(* IEC 61131-3 sources: daoli-st-library/DL_Device (part 16) *)

(* ---- FB_DL_CleanRoomRhTrim.st ---- *)
(*
  FB_DL_CleanRoomRhTrim  —  洁净室加湿阀脉冲微调（RH 偏差 + 最小开度保护） / Clean-room humidifier pulse trim with RH deviation and minimum-opening protection
  分类 Category : DL_Device
  版本 Version  : 1.0.0
  来源 Source   : t1-2-oscat-building — 楼宇洁净室湿度控制族深化
  溯源 Origin   : 道莅 clean-room 实现；脉宽调制加湿（PWM 占空比 + 最小开度 + 高限停加湿）为公开洁净室湿度算法，未复制任何源码行
  功能 Function : 1) 每个脉冲周期起始重算占空比：duty = fKpPctPerPct × (fRhSpPct - fRhPct)，
                  钳制到 [0.0, 100.0]；
                  2) 最小开度保护：fRhPct 低于 fRhLoPct 时 duty 取 max(duty, fMinOpenPct)；
                  3) 高限停加湿：fRhPct 高于 fRhHiPct 时 duty 强制 0（防过湿）；
                  4) 脉宽：开阀时长 = duty × tPeriod / 100.0（除数常量 100.0），关阀时长 = 周期余量；
                  5) 故障级单码 052B / 信息级 0431 = 脉冲周期完成沿（每周期单拍）。
  接口 Interface: 输入 RH 设定/实测/上下限/增益/最小开度/周期；输出阀指令与占空比镜像
  边界 Boundary : ① 组态闸：tPeriod <= T#0S、fMinOpenPct 不在 [0,100]、fKpPctPerPct <= 0.0、
                  fRhHiPct <= fRhLoPct、fRhSpPct 不在 [0,100] → 052B 锁存；
                  ② RH 非有限（NaN 自反 + Inf 差值自减）→ 052B 锁存，阀指令强制关断；
                  ③ 占空比开阀时长按实数乘除后转 TIME，转换前钳制到 [0, tPeriod] 防越界；
                  ④ 两个 TON 段 0 无条件周期调用，IN 由相位/占空比派生，相内自动复位 ET；
                  ⑤ 故障相迁出唯一路径 = bReset 上升沿；⑥ 零全局耦合（无 GVL / %I %Q %M）。
  依赖 Depends  : Standard.library（TON / R_TRIG）
  码表 Error codes（Device 分段见下，故障窗口 052B / 信息窗口 0431）:
    16#0003_052B 故障级：加湿脉冲故障总码（组态非法 / RH 非有限），锁存至 bReset 上升沿；
                 归因见 eCause，不新增码位（派单硬约束单码）
    16#0003_0431 信息级：脉冲周期完成沿（占空比重算单拍）
    分段理由：段 0003 故障带 03A0~03FF 于 R42 用尽，启用 05xx 副带续编，避开 0590~0599 判错位段。
  修订历史 Revision :
    2026-11-19  v1.0.0  R43 首版（批次 3 · 序号 15）
*)

TYPE E_DL_CrhState :
(
    eIdle  := 0,      // 未使能：阀关 / Idle, valve closed
    ePulse := 10,     // 脉冲调制中（开/关按时长切换） / Pulse modulation
    eFault := 90      // 故障锁存相（阀强制关） / Fault latched, valve forced closed
);
END_TYPE

TYPE E_DL_CrhCause :
(
    eNone       := 0, // 无故障成因 / No cause
    eCfgIllegal := 1, // 组态非法 / Illegal configuration
    eNonFinite  := 2  // RH 非有限 / Non-finite RH
);
END_TYPE

FUNCTION_BLOCK FB_DL_CleanRoomRhTrim
VAR_INPUT
    fRhSpPct      : REAL := 45.0;      // RH 设定 [%]，域 [0,100] / RH setpoint
    fRhPct        : REAL := 0.0;       // RH 实测 [%] / Measured RH
    fRhLoPct      : REAL := 40.0;      // 低限（触发最小开度） [%] / Low limit for minimum opening
    fRhHiPct      : REAL := 55.0;      // 高限（停加湿） [%] / High limit stopping humidification
    fKpPctPerPct  : REAL := 8.0;       // 比例增益 [%/ %]，域 > 0 / Proportional gain
    fMinOpenPct   : REAL := 10.0;      // 最小开度 [%]，域 [0,100] / Minimum opening
    tPeriod       : TIME := T#10S;     // 脉冲周期 [ms]，域 > 0 / Pulse period
    bEnable       : BOOL := FALSE;     // 加湿使能（电平）[-] / Humidification enable
    bReset        : BOOL := FALSE;     // 复位命令，上升沿清故障 [-] / Reset edge
END_VAR
VAR_OUTPUT
    eState        : E_DL_CrhState;     // 状态出口，段 6 单点映射 / State outlet
    eCause        : E_DL_CrhCause;     // 故障成因出口（R190） / Fault cause outlet
    bHumValve     : BOOL;              // 加湿阀指令 [-] / Humidifier valve command
    fDutyPct      : REAL;              // 占空比镜像 [%] / Duty mirror
    bMinOpen      : BOOL;              // 最小开度生效镜像 [-] / Minimum opening active
    bCycleDone    : BOOL;              // 脉冲周期完成标志 [-] / Pulse period done flag
    bError        : BOOL;              // 故障锁存标志 [-] / Fault latch flag
    nErrId        : UDINT;             // 事件码，0 = 无事件 / Event code
END_VAR
VAR
    _eState       : E_DL_CrhState := E_DL_CrhState.eIdle;   // 内部相位（CASE 唯一写入目标） / Internal phase
    _eCause       : E_DL_CrhCause := E_DL_CrhCause.eNone;   // 故障成因锁存（锁存量） / Latched cause
    tonOn         : TON;               // 开阀时长计时，每周期无条件调用 / Valve-on timer
    tonOff        : TON;               // 关阀时长计时，每周期无条件调用 / Valve-off timer
    rtReset       : R_TRIG;            // 复位沿实例，每周期无条件调用 / Reset edge
    _fDutyPct     : REAL;              // 占空比保持量（本周期内恒定） / Duty held for the period
    _fOnMs        : REAL;              // 本周期开阀时长 [ms]（钳制后） / On-time in ms
    _fOffMs       : REAL;              // 本周期关阀时长 [ms] / Off-time in ms
    _bOnPhase     : BOOL;              // 当前处于开阀段（内部相位标志） / In on-segment flag
    _bMinOpenOn   : BOOL;              // 最小开度生效当拍量 [-] / Minimum opening flag
    _bNonFin      : BOOL;              // RH 非有限当拍量 [-] / Non-finite RH
    _bCfgBad      : BOOL;              // 组态非法当拍量 [-] / Config illegal
    _bFault       : BOOL;              // 故障锁存位（锁存量） / Latched fault bit
    _uFault       : UDINT;             // 故障码锁存（锁存量） / Latched fault code
    _uInfo        : UDINT;             // 信息码，每拍重算 / Transient info code
END_VAR

(* —— 段 0：沿实例与定时器无条件周期刷新 + 当拍量判据 —— *)
_bNonFin := (fRhPct <> fRhPct) OR (fRhSpPct <> fRhSpPct)
         OR ((fRhPct - fRhPct) <> (fRhPct - fRhPct))
         OR ((fRhSpPct - fRhSpPct) <> (fRhSpPct - fRhSpPct));                 // NaN 自反 + Inf 差值自减 / NaN and Inf
_bCfgBad := (tPeriod <= T#0S) OR (fKpPctPerPct <= 0.0) OR (fRhHiPct <= fRhLoPct)
            OR (fMinOpenPct < 0.0) OR (fMinOpenPct > 100.0)
            OR (fRhSpPct < 0.0) OR (fRhSpPct > 100.0);                        // 组态非法当拍量 / Config illegal
rtReset(CLK := bReset);                                                       // 复位沿，每拍必调 / Reset edge
tonOn(IN := (_bOnPhase AND (_eState = E_DL_CrhState.ePulse)), PT := REAL_TO_TIME(_fOnMs));    // 开阀计时（实数时长转 TIME） / On timer
tonOff(IN := (NOT _bOnPhase) AND (_eState = E_DL_CrhState.ePulse), PT := REAL_TO_TIME(_fOffMs));  // 关阀计时 / Off timer

(* —— 段 1：单拍量预清零（锁存量与占空比保持量不入清单） —— *)
_uInfo := 16#0000_0000;            // 信息码每拍重算 / Info recomputed
bHumValve := FALSE;                // 阀指令缺省关 / Valve command default closed
fDutyPct := 0.0;                   // 占空比出口缺省 0 / Duty default
bMinOpen := FALSE;                 // 最小开度镜像缺省 FALSE / Minimum opening default
bCycleDone := FALSE;               // 周期完成标志缺省 FALSE / Period done default
nErrId := 16#0000_0000;            // 事件码缺省无事件 / Event code default

(* —— 段 2：复位沿 + 组态域闸 —— *)
IF rtReset.Q THEN                              // rtReset.Q = 当拍量 / current scan
    _bFault := FALSE;                          // 清故障锁存位（锁存量） / Clear fault latch
    _uFault := 16#0000_0000;                   // 清故障锁存码（锁存量） / Clear fault code
    _eCause := E_DL_CrhCause.eNone;            // 清成因（锁存量） / Clear cause
    _fDutyPct := 0.0;                          // 清占空比保持量 / Clear duty
    _bOnPhase := FALSE;                        // 清开阀段标志 / Clear on-segment
    IF _eState = E_DL_CrhState.eFault THEN
        _eState := E_DL_CrhState.eIdle;        // 故障相迁出：回未使能 / Fault exit to idle
    END_IF
END_IF
IF _bCfgBad THEN                               // 组态域闸 / Config gate
    _uFault := 16#0003_052B;                   // 故障级：加湿脉冲故障总码（05xx 副带） / Device fault code
    _eCause := E_DL_CrhCause.eCfgIllegal;      // 归因：组态非法 / Cause: illegal config
    _bFault := TRUE;                           // 标志与码位配对（R45） / Flag paired with code
END_IF
IF (NOT _bFault) AND _bNonFin THEN             // 非有限锁存 / Non-finite latch
    _uFault := 16#0003_052B;
    _eCause := E_DL_CrhCause.eNonFinite;       // 归因：非有限 / Cause: non-finite
    _bFault := TRUE;
END_IF

(* —— 段 3：占空比重算（周期边界 = 关阀段结束或首次进入） —— *)
IF (NOT _bFault) AND (_eState = E_DL_CrhState.ePulse) AND tonOff.Q THEN
    _fDutyPct := fKpPctPerPct * (fRhSpPct - fRhPct);                  // 比例占空比 [%] / Proportional duty
    IF fRhPct < fRhLoPct THEN                                        // 低限：最小开度保护 / Low limit protection
        IF _fDutyPct < fMinOpenPct THEN
            _fDutyPct := fMinOpenPct;                                // 抬到最小开度 / Raise to minimum
            _bMinOpenOn := TRUE;
        END_IF
    END_IF
    IF fRhPct > fRhHiPct THEN                                        // 高限：停加湿 / High limit stops humidification
        _fDutyPct := 0.0;
        _bMinOpenOn := FALSE;
    END_IF
    IF _fDutyPct < 0.0 THEN                                          // 占空比下限钳制 / Duty low clamp
        _fDutyPct := 0.0;
    ELSIF _fDutyPct > 100.0 THEN                                     // 占空比上限钳制 / Duty high clamp
        _fDutyPct := 100.0;
    END_IF
    _fOnMs := _fDutyPct / 100.0 * TIME_TO_REAL(tPeriod);             // 开阀时长 [ms]（除常量 100.0） / On-time
    IF _fOnMs < 0.0 THEN                                             // 时长下限钳制（防负数） / On-time low clamp
        _fOnMs := 0.0;
    ELSIF _fOnMs > TIME_TO_REAL(tPeriod) THEN                        // 时长上限钳制（不越周期） / On-time high clamp
        _fOnMs := TIME_TO_REAL(tPeriod);
    END_IF
    _fOffMs := TIME_TO_REAL(tPeriod) - _fOnMs;                       // 关阀时长 = 周期余量 / Off-time remainder
    _uInfo := 16#0003_0431;                                          // 信息级：脉冲周期完成沿 / Info: period done edge
END_IF

(* —— 段 4：故障解除式（R240；全当拍量）：rtReset.Q / NOT _bCfgBad / NOT _bNonFin —— *)
IF rtReset.Q AND (NOT _bCfgBad) AND (NOT _bNonFin) THEN
    _bFault := FALSE;                          // 清故障锁存位（锁存量） / Clear fault latch
    _uFault := 16#0000_0000;                   // 清故障锁存码（锁存量） / Clear fault code
    _eCause := E_DL_CrhCause.eNone;            // 清成因（锁存量） / Clear cause
END_IF

(* —— 段 4A：故障锁存相位迁移闸（阀强制关） —— *)
IF _bFault AND (_eState <> E_DL_CrhState.eFault) THEN
    _eState := E_DL_CrhState.eFault;           // 锁存即入故障相 / Latch enters fault phase
END_IF

(* —— 段 5：相位机（CASE 全覆盖 + ELSE 兜底） —— *)
CASE _eState OF

E_DL_CrhState.eIdle:
    IF bEnable AND (NOT _bFault) THEN          // 使能条件 / Enable gate
        _fDutyPct := 0.0;                      // 起始占空比 0 / Start duty zero
        _fOnMs := 0.0;                         // 起始开阀时长 0 / Start on-time zero
        _fOffMs := TIME_TO_REAL(tPeriod);      // 起始关阀时长 = 整周期 / Start off-time full period
        _bOnPhase := FALSE;                    // 从关阀段起步 / Start in off-segment
        _eState := E_DL_CrhState.ePulse;       // 进脉冲相 / Enter pulse
    END_IF

E_DL_CrhState.ePulse:
    IF _bOnPhase THEN                          // 开阀段 / On-segment
        bHumValve := TRUE;                     // 阀开 / Valve open
        IF tonOn.Q THEN                        // 开阀到时 / On-time elapsed
            _bOnPhase := FALSE;                // 转关阀段 / Switch to off-segment
        END_IF
    ELSE
        bHumValve := FALSE;                    // 阀关 / Valve closed
        IF (_fOnMs > 0.0) AND tonOff.Q THEN    // 关阀到时且有开阀时长 / Off-time elapsed with on-time
            _bOnPhase := TRUE;                 // 转开阀段 / Switch to on-segment
        ELSIF (_fOnMs <= 0.0) AND tonOff.Q THEN
            ;                                  // 零占空比：保持关阀（周期照常走完） / Zero duty keeps valve closed
            _bOnPhase := FALSE;
        END_IF
    END_IF
    IF NOT bEnable THEN                        // 撤使能：阀关，回未使能 / Disable closes valve
        _bOnPhase := FALSE;
        _eState := E_DL_CrhState.eIdle;
    END_IF

E_DL_CrhState.eFault:
    ;                                          // 故障相：阀强制关，仅段 4 复位沿可迁出 / Valve closed, reset only

ELSE
    _uFault := 16#0003_052B;                   // 故障级：非法相位兜底（归并总码） / Illegal phase fallback
    _eCause := E_DL_CrhCause.eCfgIllegal;      // 归因：相位非法归并组态 / Cause: phase illegal
    _bFault := TRUE;
    _eState := E_DL_CrhState.eFault;           // 强制回故障相 / Force fault phase

END_CASE

(* —— 段 6：出口单点映射（名实同源；故障相阀强制关断） —— *)
IF _bFault THEN
    bHumValve := FALSE;                        // 故障相阀强制关（安全侧） / Valve forced closed
    nErrId := _uFault;                         // 故障锁存码回放 / Replay latched code
    fDutyPct := 0.0;                           // 故障相占空比强制 0 / Duty forced zero
    bMinOpen := FALSE;                         // 故障相最小开度镜像强制 FALSE / Minimum opening forced false
ELSE
    nErrId := _uInfo;                          // 信息码 / Transient info
    fDutyPct := _fDutyPct;                     // 占空比镜像 / Duty mirror
    bMinOpen := _bMinOpenOn;                   // 最小开度镜像 / Minimum opening mirror
END_IF
bCycleDone := (_eState = E_DL_CrhState.ePulse) AND tonOff.Q;   // 周期完成标志（当拍量） / Period done flag
bError := _bFault;                             // 故障标志同源 / Flag from latch
eState := _eState;                             // 状态出口 / State outlet
eCause := _eCause;                             // 成因出口 / Cause outlet

END_FUNCTION_BLOCK

(* ---- FB_DL_CncLoadUnloadSeq.st ---- *)
(*
  DL Factory R84 | FB_DL_CncLoadUnloadSeq
  功能：机床上下料八相时序状态机，逐相超时置故障码并锁存至复位沿
  开源溯源：无（clean-room 自研，依据公开工艺公式，来源=行业通用公式，许可证=MIT，借鉴点=公式结构）
  规则：R1-R16 全遵守
*)
TYPE E_DL_CncUsState :
(
    eIdle := 0, // 空闲待启动 [-] / idle, waiting for start [-]
    eDoorOpen := 1, // 开门相 [-] / door opening phase [-]
    eClampOpen := 2, // 夹具松开相 [-] / clamp opening phase [-]
    ePartLoad := 3, // 上料相 [-] / part loading phase [-]
    eClampClose := 4, // 夹具夹紧相 [-] / clamp closing phase [-]
    eDoorClose := 5, // 关门相 [-] / door closing phase [-]
    eCycleStart := 6, // 加工启动相 [-] / cycle start phase [-]
    eDone := 7, // 完成相 [-] / done phase [-]
    eFault := 8 // 故障锁存相 [-] / fault latched phase [-]
) := eIdle;
END_TYPE

FUNCTION_BLOCK FB_DL_CncLoadUnloadSeq
VAR_INPUT
    xStart : BOOL; // 启动按钮 [-] / start pushbutton [-]
    xReset : BOOL; // 复位按钮（上升沿清故障码） [-] / reset pushbutton [-]
    xDoorOpened : BOOL; // 门开到位反馈 [-] / door open limit [-]
    xDoorClosed : BOOL; // 门关到位反馈 [-] / door closed limit [-]
    xClampOpened : BOOL; // 夹具松开到位反馈 [-] / clamp open limit [-]
    xClampClosed : BOOL; // 夹具夹紧到位反馈 [-] / clamp closed limit [-]
    xPartPresent : BOOL; // 工件在位检测 [-] / part present sensor [-]
    xCycleAllowed : BOOL; // 加工许可互锁（外部给定） [-] / cycle permit interlock [-]
    xCycleDone : BOOL; // 加工完成反馈 [-] / cycle finished feedback [-]
    tPhaseLimit : TIME := T#10S; // 单相超时门限 [s] / per phase timeout limit [s]
END_VAR
VAR_OUTPUT
    eState : E_DL_CncUsState; // 当前时序状态 [-] / current sequence state [-]
    iErrCode : INT; // 故障码 0=正常，101~106=逐相超时，201=非法相位 [-] / error code [-]
    xBusy : BOOL; // 时序执行中 [-] / sequence busy [-]
    xDone : BOOL; // 完成单拍脉冲 [-] / done one-shot pulse [-]
END_VAR
VAR
    rtStart : R_TRIG; // 启动上升沿实例 [-] / start rising edge instance [-]
    rtReset : R_TRIG; // 复位上升沿实例 [-] / reset rising edge instance [-]
    tonPhase : TON; // 相超时定时器（全相共用） [-] / shared phase timeout timer [-]
    xTimerRun : BOOL; // 定时器运行使能 [-] / timer run enable [-]
    tLimit : TIME; // 当前相超时设定 [s] / current phase timeout preset [s]
    xTimeout : BOOL; // 本拍超时标志 [-] / timeout flag of this scan [-]
    xDoneInt : BOOL; // 完成内部锁存位 [-] / internal done latch [-]
    xDonePrev : BOOL; // 完成前拍快照 [-] / done previous scan snapshot [-]
    _eState : E_DL_CncUsState := E_DL_CncUsState.eIdle; // 内部相位（CASE 唯一写目标） [-] / internal phase [-]
    _ePrev : E_DL_CncUsState := E_DL_CncUsState.eIdle; // 相位前拍快照（供自复位判沿） [-] / previous phase snapshot [-]
    xPhaseChg : BOOL; // 相位切换当拍标志 [-] / phase change flag of this scan [-]
    _iErr : INT; // 故障码内部锁存 [-] / latched error code [-]
END_VAR

// 段 0｜边沿实例无条件周期刷新（R7）
rtStart(CLK := xStart); // 启动沿每拍必调 [-] / start edge called every scan [-]
rtReset(CLK := xReset); // 复位沿每拍必调 [-] / reset edge called every scan [-]

// 段 1｜按相位选超时预设（必须在定时器调用之前完成）
CASE _eState OF
    E_DL_CncUsState.eIdle: tLimit := T#0S; // 空闲不计时 [s] / no timing in idle [s]
    E_DL_CncUsState.eDone: tLimit := T#0S; // 完成不计时 [s] / no timing in done [s]
    E_DL_CncUsState.eFault: tLimit := T#0S; // 故障不计时 [s] / no timing in fault [s]
ELSE
    tLimit := tPhaseLimit; // 其余工作相按门限计时 [s] / working phases use the limit [s]
END_CASE

// 段 2｜定时器无条件周期刷新（CASE 之外，无 IF 包裹；换相即自复位，R7/R188）
xPhaseChg := _eState <> _ePrev; // 相位切换沿 [-] / phase change edge [-]
xTimerRun := (((_eState <> E_DL_CncUsState.eIdle) AND (_eState <> E_DL_CncUsState.eDone)) AND (_eState <> E_DL_CncUsState.eFault)) AND NOT xPhaseChg; // 工作相定时使能，换相当拍拉低以复位计时 [-] / timing enable, dropped on a phase change to restart [-]
tonPhase(IN := xTimerRun, PT := tLimit); // 无条件刷新 [-] / unconditional refresh [-]
xTimeout := tonPhase.Q; // 本拍超时判定 [-] / timeout verdict of this scan [-]
_ePrev := _eState; // 相位快照在定时器之后更新（本拍迁移下一拍生效） [-] / phase snapshot updated after the timer call [-]

// 段 3｜复位沿：清单为故障码 + 内部锁存 + 相位，不含 Prev/Acc 保持量（R189）
IF rtReset.Q THEN
    _iErr := 0; // 清故障码 [-] / clear error code [-]
    xDoneInt := FALSE; // 清完成锁存 [-] / clear done latch [-]
    _eState := E_DL_CncUsState.eIdle; // 回空闲相 [-] / back to idle [-]
END_IF

// 段 4｜主状态机（合法事件优先于超时迁移，R275）
CASE _eState OF
    E_DL_CncUsState.eIdle: // 空闲相 [-] / idle [-]
        xDoneInt := FALSE; // 空闲清完成锁存 [-] / clear done latch in idle [-]
        IF rtStart.Q THEN
            _eState := E_DL_CncUsState.eDoorOpen; // 启动沿开安全门 [-] / start edge opens the door [-]
        END_IF
    E_DL_CncUsState.eDoorOpen: // 开门相 [-] / door opening [-]
        IF xDoorOpened THEN
            _eState := E_DL_CncUsState.eClampOpen; // 门开到位转松夹 [-] / door open leads to clamp open [-]
        ELSIF xTimeout THEN
            _iErr := 101; _eState := E_DL_CncUsState.eFault; // 开门超时 [-] / door open timeout [-]
        END_IF
    E_DL_CncUsState.eClampOpen: // 松夹相 [-] / clamp opening [-]
        IF xClampOpened THEN
            _eState := E_DL_CncUsState.ePartLoad; // 松夹到位转上料 [-] / clamp open leads to loading [-]
        ELSIF xTimeout THEN
            _iErr := 102; _eState := E_DL_CncUsState.eFault; // 松夹超时 [-] / clamp open timeout [-]
        END_IF
    E_DL_CncUsState.ePartLoad: // 上料相 [-] / part loading [-]
        IF xPartPresent AND NOT xTimeout THEN
            _eState := E_DL_CncUsState.eClampClose; // 工件在位转夹紧（带超时复检） [-] / part present leads to clamp close [-]
        ELSIF xTimeout THEN
            _iErr := 103; _eState := E_DL_CncUsState.eFault; // 上料超时（工件未到位） [-] / loading timeout [-]
        END_IF
    E_DL_CncUsState.eClampClose: // 夹紧相 [-] / clamp closing [-]
        IF xClampClosed THEN
            _eState := E_DL_CncUsState.eDoorClose; // 夹紧到位转关门 [-] / clamp closed leads to door close [-]
        ELSIF xTimeout THEN
            _iErr := 104; _eState := E_DL_CncUsState.eFault; // 夹紧超时 [-] / clamp close timeout [-]
        END_IF
    E_DL_CncUsState.eDoorClose: // 关门相 [-] / door closing [-]
        IF xDoorClosed THEN
            _eState := E_DL_CncUsState.eCycleStart; // 关门到位转加工启动 [-] / door closed leads to cycle start [-]
        ELSIF xTimeout THEN
            _iErr := 105; _eState := E_DL_CncUsState.eFault; // 关门超时 [-] / door close timeout [-]
        END_IF
    E_DL_CncUsState.eCycleStart: // 加工启动相（执行类安全相，入相全量复检） [-] / cycle start [-]
        IF xCycleDone THEN
            _eState := E_DL_CncUsState.eDone; // 加工完成转完成相 [-] / cycle done leads to done [-]
        ELSIF NOT (xCycleAllowed AND xDoorClosed) THEN
            _iErr := 106; _eState := E_DL_CncUsState.eFault; // 许可消失即故障（不空等） [-] / permit lost becomes fault [-]
        ELSIF xTimeout THEN
            _iErr := 106; _eState := E_DL_CncUsState.eFault; // 加工未完成超时 [-] / cycle start timeout [-]
        END_IF
    E_DL_CncUsState.eDone: // 完成相 [-] / done [-]
        xDoneInt := TRUE; // 置完成锁存（出口统一映射单拍） [-] / raise done latch [-]
        IF NOT xStart THEN
            _eState := E_DL_CncUsState.eIdle; // 松开启动即回空闲 [-] / start released returns to idle [-]
        END_IF
    E_DL_CncUsState.eFault: // 故障相：码值锁存回放，仅复位沿出 [-] / fault, exit only on reset edge [-]
        ; // 锁存回放，不按当下输入重新推断（R28） [-] / replay the latch only [-]
ELSE
    _iErr := 201; _eState := E_DL_CncUsState.eFault; // 非法相位兜底 [-] / illegal phase fallback [-]
END_CASE

// 段 5｜出口映射（名实双出口，同源赋值）
eState := _eState; // 状态出口 [-] / state outlet [-]
iErrCode := _iErr; // 故障码出口（锁存值） [-] / error code outlet [-]
xBusy := ((_eState <> E_DL_CncUsState.eIdle) AND (_eState <> E_DL_CncUsState.eDone)) AND (_eState <> E_DL_CncUsState.eFault); // 忙 = 工作相镜像 [-] / busy mirrors a working phase [-]
xDone := xDoneInt AND NOT xDonePrev; // 完成单拍（内部锁存 → 出口映射） [-] / done one-shot [-]
xDonePrev := xDoneInt; // 本拍快照供下拍比较 [-] / snapshot for the next scan [-]
END_FUNCTION_BLOCK

(* ---- FB_DL_CncToolWearCompLoop.st ---- *)
(*
  DL Factory R84 | FB_DL_CncToolWearCompLoop
  功能：CNC 刀具后刀面磨损量 VB 在线估计与刀补闭环：按切削路程三段线性磨损曲线出 VB 原值，按切削比能调制滤波增益做一阶指数平滑得 VB 估计，超补偿门限按增量限幅出刀补，超寿命锁存换刀请求。
  开源溯源：无（clean-room 自研，依据公开工艺公式与安全设计惯例，来源=行业通用公式+工程实践，许可证=MIT，借鉴点=公式结构与联锁分层）
  规则：R1-R16 全遵守
  ------------------------------------------------------------------
  分类 DL_Device ｜ 复杂度 cx4 ｜ 版本 v1.0.0 ｜ 平台 纯 IEC 61131-3（LREAL、ENUM、CASE）
  边界一：只出刀补增量与换刀请求，不驱动伺服轴、不写 CNC 刀补表（落表由上层 PRG 执行，属主边界）。
  边界二：磨损曲线为三段线性——初期占额定寿命路程 0.15 段、占磨损余量 0.30 份；稳态占 0.70 段、占 0.55 份；
          急剧占余下 0.15 段、占余下 0.15 份；三段积分在路程等于额定寿命处恰等于 VB 限值（量纲自检见下）。
  边界三：切削路程按「进给率 × 切削时长增量」积分，时长增量取 fCutTimeS 的上拍快照差分（R45 ②）；
          负增量判零、超大跳变钳到 1 秒，防掉电恢复的时钟跳变伪造路程。
  边界四：工艺代理常量——DL_CNC_AP_MM 与 DL_CNC_AE_MM 为名义切深与切宽代理值（本件无切深切宽引脚）；
          代理值是名义切深切宽、覆盖常规铣削 0.2~3 mm 切深与 4~20 mm 切宽区间、区间外的重型切槽工况由上层
          按实际切深切宽折算 fKcNmm2 后下发（R95 三句齐备，代理假设挂编译验证债）。
  边界五：无效拍语义——功率或转速为零、或任一浮点入参非有限 → xValid 出假、相位保持、刀补增量出零；
          不推进滤波、不累加路程（不除零、不外推）。
  边界六：换刀请求 xChangeReq 为锁存式，唯一解除路径为 bReset 上升沿（R188）；xAlarm 为电平式跟随相位。
  量纲自检：VB [mm]＝斜率 [mm/m] × 路程 [m]；斜率一 ＝ VB限值 × 0.30 ÷（额定寿命 × 0.15）[mm/m]；
          路程增量 [m]＝进给 [mm/min] × 时长增量 [s] ÷ 60 [s/min] × 0.001 [m/mm]；
          切削功率 [kW]＝Kc [N/mm²] × 切除率 [mm³/s] ÷ 1000 [W/kW]；
          切除率 [mm³/s]＝进给 [mm/s] × 切深 [mm] × 切宽 [mm]；刀补 [µm]＝VB [mm] × 1000 [µm/mm]。
  码表：本件全部码位为信息级（2601 非法相位、2602 组态越域、2603 入参非有限、2604 转速或功率为零）；
        信息级码每拍重算且不置 bError；故障级语义由 xChangeReq 锁存位承担，故本件无 bError 出口（R187）。
  输出契约：fCompUm 为本次刀补增量 [µm]（限幅 ±50，非补偿相出 0 不保持）；fCompAccUm 为累计刀补 [µm]（0~200 单向）；
          fVbEst 为滤波后估计 [mm]；fVbRaw 为曲线原值 [mm]；iErrCode 信息级，非零时 xValid 恒假。
  修订记录：2026-11-24 v1.0.0 R84 首版（批 R84 · 序号 41）
*)

TYPE E_DL_CncWearState :
(
    eIdle       := 0,  // 空闲：等使能与切削条件 / idle, waiting for the enable and the cutting condition
    eLearn      := 10, // 学习：累加路程并收敛 VB 滤波 / learning, accumulate the path and settle the filter
    eCompensate := 20, // 补偿：VB 超补偿门限，按增量出刀补 / compensating, the wear passed the trigger threshold
    eAlarm      := 30, // 报警：VB 超报警门限，继续补偿并报警 / alarm, the wear passed the alarm threshold
    eChangeReq  := 40  // 换刀请求：VB 超寿命，锁存至复位沿 / change request, the wear passed the life limit and is latched
);
END_TYPE

TYPE E_DL_CncWearCause :
(
    eNone      := 0, // 无成因 / no cause
    ePhaseBad  := 1, // 非法相位（信息级 2601）/ illegal phase, info grade 2601
    eCfgBad    := 2, // 组态越域（信息级 2602）/ the configuration is out of its domain, info grade 2602
    eNotFinite := 3, // 入参非有限（信息级 2603）/ a non-finite input, info grade 2603
    eSpeedZero := 4  // 转速或功率为零（信息级 2604）/ the speed or the power is zero, info grade 2604
);
END_TYPE

FUNCTION_BLOCK FB_DL_CncToolWearCompLoop
VAR CONSTANT
    DL_CNC_PH1_FRAC   : LREAL := 0.15;    // 初期磨损段占额定寿命的路程分数 [-] / the initial wear path fraction of the rated life [-]
    DL_CNC_PH1_WEAR   : LREAL := 0.30;    // 初期磨损段占磨损余量的份额 [-] / the initial wear share of the allowance [-]
    DL_CNC_PH2_FRAC   : LREAL := 0.70;    // 稳态磨损段占额定寿命的路程分数 [-] / the steady wear path fraction of the rated life [-]
    DL_CNC_PH2_WEAR   : LREAL := 0.55;    // 稳态磨损段占磨损余量的份额 [-] / the steady wear share of the allowance [-]
    DL_CNC_ALARM_FRAC : LREAL := 0.85;    // 报警门限回退系数（组态越域时用）[-] / the alarm threshold fallback factor [-]
    DL_CNC_HYST_BAND  : LREAL := 0.02;    // 报警相回补偿相的回差带（VB 限值倍数）[-] / the hysteresis band for the alarm exit [-]
    DL_CNC_ALPHA_MIN  : LREAL := 0.02;    // 滤波增益下限（防迟钝）[-] / the filter gain lower bound [-]
    DL_CNC_ALPHA_MAX  : LREAL := 0.50;    // 滤波增益上限（防抖动）[-] / the filter gain upper bound [-]
    DL_CNC_ALPHA_SPAN : LREAL := 0.50;    // 比能超出量归一跨度（比能比 - 1 的满量程）[-] / the normalised span of the specific energy excess [-]
    DL_CNC_PWR_GAIN   : LREAL := 0.80;    // 比能超基准对磨损的加速增益 [-] / the specific energy excess gain on the wear [-]
    DL_CNC_ACCEL_MAX  : LREAL := 3.00;    // 加速因子上限 [-] / the acceleration factor upper bound [-]
    DL_CNC_RATIO_BAND : LREAL := 0.02;    // 比能比值的容差带（浮点比较）[-] / the specific energy ratio tolerance band [-]
    DL_CNC_VB_HEAD    : LREAL := 2.00;    // VB 估计上限（VB 限值倍数，防过冲）[-] / the VB estimate headroom over the limit [-]
    DL_CNC_STEP_UM    : LREAL := 50.0;    // 单次刀补增量限幅 [µm] / the per-scan compensation step limit [um]
    DL_CNC_ACC_UM     : LREAL := 200.0;   // 累计刀补上限 [µm] / the accumulated compensation upper limit [um]
    DL_CNC_UM_PER_MM  : LREAL := 1000.0;  // 毫米到微米折算系数 [µm/mm] / the millimetre to micrometre factor [um/mm]
    DL_CNC_M_PER_MM   : LREAL := 0.001;   // 毫米到米折算系数 [m/mm] / the millimetre to metre factor [m/mm]
    DL_CNC_SEC_MIN    : LREAL := 60.0;    // 秒到分钟折算系数 [s/min] / the second to minute factor [s/min]
    DL_CNC_W_PER_KW   : LREAL := 1000.0;  // 瓦到千瓦折算系数 [W/kW] / the watt to kilowatt factor [W/kW]
    DL_CNC_DTJUMP_S   : LREAL := 1.0;     // 切削时长增量上限（时钟跳变钳位）[s] / the cutting time increment upper clamp [s]
    DL_CNC_AP_MM       : LREAL := 1.0;    // 名义轴向切深代理值 [mm] / the nominal axial depth of cut proxy [mm]
    DL_CNC_AE_MM       : LREAL := 10.0;   // 名义径向切宽代理值 [mm] / the nominal radial width of cut proxy [mm]
    DL_CNC_EPS         : LREAL := 1.0E-9; // 除法零闸与零判定门限 [-] / the division guard and zero test threshold [-]
END_VAR
VAR_INPUT
    bEnable        : BOOL := TRUE;    // 使能，失能回空闲且刀补增量归零 [-] / enable, a disable returns to idle with the step zeroed
    bReset         : BOOL := FALSE;   // 复位上升沿清换刀请求锁存 [-] / reset rising edge clears the change request latch
    bCutting       : BOOL := FALSE;   // 切削中，为真才累加切削路程 [-] / cutting active, the path accumulates only while true
    fSpindleKw     : LREAL := 0.0;    // 主轴有功功率 [kW] / the spindle active power [kW]
    fFeedMmMin     : LREAL := 0.0;    // 进给率 [mm/min] / the feed rate [mm/min]
    fRpm           : LREAL := 0.0;    // 主轴转速 [r/min] / the spindle speed [r/min]
    fCutTimeS      : LREAL := 0.0;    // 本刀具累计切削时长（由上层保持）[s] / the accumulated cutting time of the tool [s]
    fKcNmm2        : LREAL := 2000.0; // 材料单位切削力系数 [N/mm²] / the specific cutting force coefficient [N/mm^2]
    fVbLimitMm     : LREAL := 0.30;   // 后刀面磨损量限值（换刀门限）[mm] / the flank wear limit, the change threshold [mm]
    fLifePathM     : LREAL := 8000.0; // 刀具额定寿命切削路程 [m] / the rated cutting path of the tool life [m]
    fIdleKw        : LREAL := 0.5;    // 主轴空载功率（扣除项）[kW] / the spindle idle power to be deducted [kW]
    fVbCompTrigMm  : LREAL := 0.15;   // 补偿启动门限 [mm] / the compensation trigger threshold [mm]
    fVbAlarmMm     : LREAL := 0.25;   // 报警门限 [mm] / the alarm threshold [mm]
END_VAR
VAR_OUTPUT
    fVbEst      : LREAL := 0.0;   // 滤波后磨损量估计 [mm] / the filtered wear estimate [mm]
    fVbRaw      : LREAL := 0.0;   // 磨损曲线原值（未滤波）[mm] / the raw wear from the piecewise curve [mm]
    fCompUm     : LREAL := 0.0;   // 本次刀补增量 [µm] / the compensation increment of this scan [um]
    fCompAccUm  : LREAL := 0.0;   // 累计刀补量 [µm] / the accumulated compensation [um]
    fPathM      : LREAL := 0.0;   // 累计切削路程 [m] / the accumulated cutting path [m]
    fKcRatio    : LREAL := 1.0;   // 实测比能比（切削功率 ÷ 名义切削功率）[-] / the measured specific energy ratio [-]
    xChangeReq  : BOOL := FALSE;  // 换刀请求（锁存式，复位沿清除）[-] / the change request, latched until the reset edge
    xAlarm      : BOOL := FALSE;  // 磨损报警（电平式）[-] / the wear alarm, level type
    eState      : E_DL_CncWearState := E_DL_CncWearState.eIdle; // 相位出口 [枚举] / the phase outlet [enum]
    iErrCode    : INT := 0;       // 信息级码（每拍重算，非锁存）[码] / the info grade code, recomputed every scan [code]
    xValid      : BOOL := FALSE;  // 本拍估计可信（判据全通过）[-] / the estimate is trustworthy this scan [-]
END_VAR
VAR
    rtReset : R_TRIG; // 复位上升沿实例（R188：电平复位会导致按住即反复清零） [-] / reset rising edge instance [-]
    _eState     : E_DL_CncWearState := E_DL_CncWearState.eIdle; // 内部相位（枚举，无量纲）[-] / the internal phase, the only CASE target
    _bInit      : BOOL := FALSE;  // 首扫初始化完成标志（R310）[-] / the first scan initialisation flag [-]
    _bFinOk     : BOOL := FALSE;  // 全部浮点入参有限 [-] / every floating input is finite
    _bCfgOk     : BOOL := FALSE;  // 组态参数域内 [-] / the configuration is inside its domain
    _bSpeedOk   : BOOL := FALSE;  // 转速与功率非零（防除零）[-] / the speed and the power are non zero
    _bValid     : BOOL := FALSE;  // 三个闸的合取 [-] / the conjunction of the three gates
    _bChangeLch : BOOL := FALSE;  // 换刀请求锁存位（唯一清除：复位沿）[-] / the change request latch, cleared by the reset edge only
    _iErrTmp    : INT := 0;       // 本拍信息级码暂存 [码] / the scan info code scratch [code]
    _fCutPrevS  : LREAL := 0.0;   // 上拍切削时长快照（差分用）[s] / the previous scan cutting time snapshot [s]
    _fDtCutS    : LREAL := 0.0;   // 切削时长增量（钳定后）[s] / the clamped cutting time increment [s]
    _fPathM     : LREAL := 0.0;   // 累计切削路程（跨批保持）[m] / the accumulated cutting path across batches [m]
    _fPnomKw    : LREAL := 0.0;   // 名义切削功率 [kW] / the nominal cutting power [kW]
    _fPcKw      : LREAL := 0.0;   // 实测净切削功率（扣除空载）[kW] / the measured net cutting power [kW]
    _fRatio     : LREAL := 1.0;   // 比能比（含域夹取）[-] / the specific energy ratio with clamping [-]
    _fExcess    : LREAL := 0.0;   // 比能超出量归一值 [0,1] [-] / the normalised specific energy excess [-]
    _fAlpha     : LREAL := 0.0;   // 本拍滤波增益（随比能自适应）[-] / the adaptive filter gain of this scan [-]
    _fSlope1    : LREAL := 0.0;   // 初期磨损段斜率 [mm/m] / the initial wear slope [mm/m]
    _fSlope2    : LREAL := 0.0;   // 稳态磨损段斜率 [mm/m] / the steady wear slope [mm/m]
    _fSlope3    : LREAL := 0.0;   // 急剧磨损段斜率 [mm/m] / the severe wear slope [mm/m]
    _fL1        : LREAL := 0.0;   // 初期磨损段终点路程 [m] / the initial wear segment end path [m]
    _fL2        : LREAL := 0.0;   // 稳态磨损段终点路程 [m] / the steady wear segment end path [m]
    _fAccel     : LREAL := 1.0;   // 比能加速因子 [-] / the specific energy acceleration factor [-]
    _fVbRaw     : LREAL := 0.0;   // 磨损曲线原值 [-] / the raw wear value [-]
    _fVbFilt    : LREAL := 0.0;   // 滤波后磨损量（保持槽，写入前过非有限闸）[mm] / the filtered wear, guarded before the write [mm]
    _fVbEst     : LREAL := 0.0;   // 本拍磨损估计 [mm] / the wear estimate of this scan [mm]
    _fAlarmMm   : LREAL := 0.0;   // 报警门限（两级回退后）[mm] / the alarm threshold after the two level fallback [mm]
    _fCompAcc   : LREAL := 0.0;   // 累计刀补量 [µm] / the accumulated compensation [um]
    _fCompTgt   : LREAL := 0.0;   // 目标累计刀补量 [µm] / the target accumulated compensation [um]
    _fStep      : LREAL := 0.0;   // 本拍刀补增量（限幅后）[µm] / the limited compensation step of this scan [um]
END_VAR
// 段 0｜出口预置：所有出口先赋安全侧值，任何早退路径不留未初始化输出
xValid := FALSE; // 有效性预置假（判据未完成前一律无效，安全侧）/ validity preset false on the safe side
xAlarm := FALSE; // 报警预置假 / the alarm preset false
xChangeReq := _bChangeLch; // 换刀请求回放锁存位 / replay the change request latch
fCompUm := 0.0; // 刀补增量预置零（非补偿相不出量）/ the step preset zero while not compensating
fVbEst := 0.0; // 估计预置零 / the estimate preset zero
fVbRaw := 0.0; // 原值预置零 / the raw value preset zero
fCompAccUm := _fCompAcc; // 累计刀补回放 / replay the accumulated compensation
fPathM := _fPathM; // 路程回放 / replay the path
fKcRatio := _fRatio; // 比能比回放 / replay the specific energy ratio
eState := _eState; // 相位回放 / replay the phase
iErrCode := 0; // 信息级码预置零（本拍重算）/ the info code preset zero, recomputed this scan
_iErrTmp := 0; // 单拍码暂存预清零（FB32-1：仅单拍标志可预清）/ preclear the scan code scratch only
// 段 1｜非有限闸：NaN 用自反比较、Inf 用差值自减双判，逐项枚举全部浮点入参（R79、R272）
_bFinOk := (fSpindleKw = fSpindleKw) AND ((fSpindleKw - fSpindleKw) = (fSpindleKw - fSpindleKw)) // 主轴功率有限 [-] / the spindle power is finite
    AND (fFeedMmMin = fFeedMmMin) AND ((fFeedMmMin - fFeedMmMin) = (fFeedMmMin - fFeedMmMin)) // 进给率有限 [-] / the feed rate is finite
    AND (fRpm = fRpm) AND ((fRpm - fRpm) = (fRpm - fRpm)) // 转速有限 [-] / the speed is finite
    AND (fCutTimeS = fCutTimeS) AND ((fCutTimeS - fCutTimeS) = (fCutTimeS - fCutTimeS)) // 切削时长有限 [-] / the cutting time is finite
    AND (fKcNmm2 = fKcNmm2) AND ((fKcNmm2 - fKcNmm2) = (fKcNmm2 - fKcNmm2)) // 切削力系数有限 [-] / the cutting force coefficient is finite
    AND (fVbLimitMm = fVbLimitMm) AND ((fVbLimitMm - fVbLimitMm) = (fVbLimitMm - fVbLimitMm)) // 磨损限值有限 [-] / the wear limit is finite
    AND (fLifePathM = fLifePathM) AND ((fLifePathM - fLifePathM) = (fLifePathM - fLifePathM)) // 额定寿命路程有限 [-] / the rated life path is finite
    AND (fIdleKw = fIdleKw) AND ((fIdleKw - fIdleKw) = (fIdleKw - fIdleKw)) // 空载功率有限 [-] / the idle power is finite
    AND (fVbCompTrigMm = fVbCompTrigMm) AND ((fVbCompTrigMm - fVbCompTrigMm) = (fVbCompTrigMm - fVbCompTrigMm)) // 补偿门限有限 [-] / the trigger threshold is finite
    AND (fVbAlarmMm = fVbAlarmMm) AND ((fVbAlarmMm - fVbAlarmMm) = (fVbAlarmMm - fVbAlarmMm)); // 报警门限有限 [-] / the alarm threshold is finite
// 段 2｜组态域闸：门限次序与正定性，参与判据换算的每个引脚都在闸内（R151）
_bCfgOk := (fVbLimitMm > 0.0) AND (fLifePathM > 0.0) AND (fKcNmm2 > 0.0) AND (fIdleKw >= 0.0) // 限值、寿命、系数、空载功率四项域闸 [-] / the four base domains
    AND (fVbCompTrigMm > 0.0) AND (fVbCompTrigMm < fVbLimitMm) // 补偿门限介于零与限值之间 [-] / the trigger sits between zero and the limit
    AND (fVbAlarmMm > fVbCompTrigMm) AND (fVbAlarmMm <= fVbLimitMm); // 报警门限高于补偿门限且不超限值 [-] / the alarm sits above the trigger and never above the limit
_bSpeedOk := (ABS(fRpm) > DL_CNC_EPS) AND (ABS(fSpindleKw) > DL_CNC_EPS); // 转速与功率非零闸（防除零，R4）/ the non zero gate against the division by zero
_bValid := _bFinOk AND _bCfgOk AND _bSpeedOk; // 三个闸合取 / the conjunction of the three gates
IF NOT _bFinOk THEN _iErrTmp := 2603; ELSIF NOT _bCfgOk THEN _iErrTmp := 2602; ELSIF NOT _bSpeedOk THEN _iErrTmp := 2604; END_IF // 信息级码分派（有限 → 组态 → 零速）/ the info code dispatch
// 段 3｜首扫初始化与复位沿同块，作用域逐项声明（R310、R311）
rtReset(CLK := bReset); // 复位沿无条件周期刷新（R7） [-] / the reset edge refreshed every scan [-]

IF (NOT _bInit) OR rtReset.Q THEN // 首扫一拍或复位上升沿（R188，禁电平复位） / the first scan or the reset edge
    _bInit := TRUE; // 首扫完成标志（复位沿重复置位同效）/ the first scan flag, the same effect on reset
    _bChangeLch := FALSE; // 作用域一：清换刀请求锁存（唯一清除边，R188）/ scope one, clear the change request latch
    _fVbFilt := 0.0; // 作用域二：清滤波保持槽 / scope two, clear the filter hold slot
    _fCompAcc := 0.0; // 作用域二：清累计刀补 / scope two, clear the accumulated compensation
    _fPathM := 0.0; // 作用域三：清切削路程（换刀后按新刀重计）/ scope three, clear the path for the new tool
    _fCutPrevS := fCutTimeS; // 作用域三：时长快照重取（防跨批假路程）/ scope three, re-take the snapshot
    _eState := E_DL_CncWearState.eIdle; // 作用域二：迁回空闲相 / scope two, migrate to idle
END_IF
// 段 4｜切削路程积分：时长增量差分 + 双向钳定，仅有效拍且切削中累加（R45 ②）
_fDtCutS := fCutTimeS - _fCutPrevS; // 切削时长增量 [s] / the cutting time increment [s]
IF _fDtCutS < 0.0 THEN _fDtCutS := 0.0; END_IF // 负增量判零（时钟回退不伪造路程）/ a negative increment is zeroed
IF _fDtCutS > DL_CNC_DTJUMP_S THEN _fDtCutS := DL_CNC_DTJUMP_S; END_IF // 超大跳变钳位（掉电恢复不伪造路程）/ a huge jump is clamped
IF _bValid AND bCutting THEN // 仅有效拍且切削中 / only on a valid scan while cutting
    _fPathM := _fPathM + fFeedMmMin * (_fDtCutS / DL_CNC_SEC_MIN) * DL_CNC_M_PER_MM; // 路程增量 [m] / the path increment [m]
END_IF
_fCutPrevS := fCutTimeS; // 上拍时长快照（用完立即赋值，防重复累计）/ the snapshot taken right after the integration
// 段 5｜切削比能：名义功率由 Kc 与名义切除率折算（切深切宽取边界四之代理常量），分母显式零闸（R4）
IF _bValid THEN // 仅在有效拍计算比能 / compute the ratio on a valid scan only
    _fPnomKw := fKcNmm2 * (fFeedMmMin / DL_CNC_SEC_MIN) * DL_CNC_AP_MM * DL_CNC_AE_MM / (DL_CNC_W_PER_KW * 1000.0); // N/mm2·mm3/s = mW，再除以 1e6 得 kW（量纲校正，R583） / [N/mm2]*[mm3/s] = [mW], divided by 1e6 for [kW]
    _fPcKw := fSpindleKw - fIdleKw; // 净切削功率 [kW] / the net cutting power [kW]
    IF _fPcKw < 0.0 THEN _fPcKw := 0.0; END_IF // 负净功率夹取（空载波动）/ clamp the negative net power
    _fRatio := 1.0; // 比能比默认一（无切除按名义）/ the ratio defaults to one without stock removal
    IF (_fPnomKw > DL_CNC_EPS) AND (fFeedMmMin > DL_CNC_EPS) THEN // 双分母零闸 / both denominators guarded
        _fRatio := _fPcKw / _fPnomKw; // 比能比 [-] / the specific energy ratio [-]
    END_IF
    IF _fRatio < 0.2 THEN _fRatio := 0.2; ELSIF _fRatio > 3.0 THEN _fRatio := 3.0; END_IF // 比值域夹取，防加速因子发散 / clamp the ratio domain
END_IF
// 段 6｜三段线性磨损曲线：三段斜率由额定寿命与 VB 限值反算，积分在寿命终点恰为限值
IF _bCfgOk THEN // 组态域内才反算斜率（分母中含 fLifePathM，越域即除零）/ compute the slopes only inside the domain
    _fSlope1 := (fVbLimitMm * DL_CNC_PH1_WEAR) / (fLifePathM * DL_CNC_PH1_FRAC); // 初期段斜率 [mm/m] / the initial slope [mm/m]
    _fSlope2 := (fVbLimitMm * DL_CNC_PH2_WEAR) / (fLifePathM * DL_CNC_PH2_FRAC); // 稳态段斜率 [mm/m] / the steady slope [mm/m]
    _fSlope3 := (fVbLimitMm * (1.0 - DL_CNC_PH1_WEAR - DL_CNC_PH2_WEAR)) / (fLifePathM * (1.0 - DL_CNC_PH1_FRAC - DL_CNC_PH2_FRAC)); // 急剧段斜率 [mm/m] / the severe slope [mm/m]
    _fL1 := fLifePathM * DL_CNC_PH1_FRAC; // 初期段终点 [m] / the initial segment end [m]
    _fL2 := _fL1 + fLifePathM * DL_CNC_PH2_FRAC; // 稳态段终点 [m] / the steady segment end [m]
    IF _fPathM <= _fL1 THEN // 阶段一：初期磨损 / stage one, the initial wear
        _fVbRaw := _fSlope1 * _fPathM; // 初期段磨损 [mm] / the initial wear [mm]
    ELSIF _fPathM <= _fL2 THEN // 阶段二：稳态磨损（含初期段积分）/ stage two, the steady wear including the initial integral
        _fVbRaw := _fSlope1 * _fL1 + _fSlope2 * (_fPathM - _fL1); // 稳态段磨损 [mm] / the steady wear [mm]
    ELSE // 阶段三：急剧磨损 / stage three, the severe wear
        _fVbRaw := _fSlope1 * _fL1 + _fSlope2 * (_fL2 - _fL1) + _fSlope3 * (_fPathM - _fL2); // 急剧段磨损 [mm] / the severe wear [mm]
    END_IF
    IF _fRatio > (1.0 + DL_CNC_RATIO_BAND) THEN // 比能高于基准才加速 / accelerate only above the base
        _fAccel := 1.0 + DL_CNC_PWR_GAIN * (_fRatio - 1.0); // 加速因子 [-] / the acceleration factor [-]
    ELSE // 比能未超基准：不加速也不抑制 / no acceleration below the base
        _fAccel := 1.0; // 加速因子归一 / the factor is unity
    END_IF
    IF _fAccel > DL_CNC_ACCEL_MAX THEN _fAccel := DL_CNC_ACCEL_MAX; END_IF // 加速因子上限 / the factor upper bound
    _fVbRaw := _fVbRaw * _fAccel; // 比能修正后磨损 [mm] / the wear corrected by the specific energy
    IF _fVbRaw > (fVbLimitMm * DL_CNC_VB_HEAD) THEN _fVbRaw := fVbLimitMm * DL_CNC_VB_HEAD; END_IF // 上限兜底防过冲 / the upper bound against overshoot
END_IF
// 段 7｜一阶指数滤波：增益随比能超出量自适应（钝化加剧时跟随更快），写入前过非有限闸（R133）
_fExcess := (_fRatio - 1.0) / DL_CNC_ALPHA_SPAN; // 超出量归一 [-] / the normalised excess [-]
IF _fExcess < 0.0 THEN _fExcess := 0.0; ELSIF _fExcess > 1.0 THEN _fExcess := 1.0; END_IF // 归一值夹取到 [0,1] / clamp the excess into [0,1]
_fAlpha := DL_CNC_ALPHA_MIN + (DL_CNC_ALPHA_MAX - DL_CNC_ALPHA_MIN) * _fExcess; // 本拍增益 [-] / the gain of this scan [-]
IF _bValid THEN // 仅有效拍推进滤波（无效拍不污染保持槽）/ advance only on a valid scan
    _fVbFilt := _fVbFilt + _fAlpha * (_fVbRaw - _fVbFilt); // 一阶指数平滑 [mm] / the first order exponential smoothing [mm]
END_IF
IF NOT (_fVbFilt = _fVbFilt) THEN _fVbFilt := _fVbRaw; END_IF // 滤波结果 NaN 兜底（回退原值）/ the NaN fallback to the raw value
IF (_fVbFilt - _fVbFilt) <> (_fVbFilt - _fVbFilt) THEN _fVbFilt := _fVbRaw; END_IF // 滤波结果 Inf 兜底（同回退）/ the Inf fallback to the raw value
_fVbEst := _fVbFilt; // 本拍估计 [mm] / the estimate of this scan [mm]
IF _fVbEst < 0.0 THEN _fVbEst := 0.0; END_IF // 估计下限夹取（磨损不可为负）/ the wear can never be negative
// 段 8｜报警门限两级回退：一级回默认系数、二级按有效域钳定（R117）
_fAlarmMm := fVbAlarmMm; // 一级：取引脚值 / level one, take the pin value
IF NOT _bCfgOk THEN // 组态越域：一级回退到限值系数 / out of domain, fall back to the limit factor
    _fAlarmMm := fVbLimitMm * DL_CNC_ALARM_FRAC; // 回退值 [mm] / the fallback threshold [mm]
    IF _fAlarmMm <= fVbCompTrigMm THEN _fAlarmMm := fVbCompTrigMm + (fVbLimitMm * DL_CNC_RATIO_BAND); END_IF // 二级：按有效域钳定 / level two, clamp into the valid domain
END_IF
// 段 9｜相位状态机：ENUM ＋ CASE ＋ ELSE 非法相位兜底（R6、R128）
CASE _eState OF
E_DL_CncWearState.eIdle: // 空闲相：退出条件三（使能、切削中、有效拍、无换刀锁存）
    IF _bChangeLch THEN // 换刀请求未解除：禁止回到生产 / the change request blocks production
        _eState := E_DL_CncWearState.eChangeReq; // 驻留换刀请求相 / stay in the change request phase
    ELSIF bEnable AND bCutting AND _bValid THEN // 三个条件齐备才进学习 / all three conditions enter learning
        _eState := E_DL_CncWearState.eLearn; // 迁学习相 / migrate to learning
    END_IF
E_DL_CncWearState.eLearn: // 学习相：按门限升相，无门限命中则驻留（驻留由注释表达，禁自赋值 R261）
    IF NOT bEnable THEN // 使能丢失 / the enable was lost
        _eState := E_DL_CncWearState.eIdle; // 回空闲 / back to idle
    ELSIF _fVbEst >= fVbLimitMm THEN // 越过寿命限值 / the life limit was passed
        _eState := E_DL_CncWearState.eChangeReq; // 迁换刀请求相 / migrate to the change request
    ELSIF _fVbEst >= _fAlarmMm THEN // 越过报警门限 / the alarm threshold was passed
        _eState := E_DL_CncWearState.eAlarm; // 迁报警相 / migrate to alarm
    ELSIF _fVbEst >= fVbCompTrigMm THEN // 越过补偿门限 / the trigger threshold was passed
        _eState := E_DL_CncWearState.eCompensate; // 迁补偿相 / migrate to compensating
    END_IF
E_DL_CncWearState.eCompensate: // 补偿相：按门限升相，回落到补偿门限以下不降相（已补量不回退）
    IF NOT bEnable THEN // 使能丢失 / the enable was lost
        _eState := E_DL_CncWearState.eIdle; // 回空闲 / back to idle
    ELSIF _fVbEst >= fVbLimitMm THEN // 越过寿命限值 / the life limit was passed
        _eState := E_DL_CncWearState.eChangeReq; // 迁换刀请求相 / migrate to the change request
    ELSIF _fVbEst >= _fAlarmMm THEN // 越过报警门限 / the alarm threshold was passed
        _eState := E_DL_CncWearState.eAlarm; // 迁报警相 / migrate to alarm
    END_IF
E_DL_CncWearState.eAlarm: // 报警相：退出条件三（使能丢失、升换刀、带回差降回补偿）
    IF NOT bEnable THEN // 使能丢失 / the enable was lost
        _eState := E_DL_CncWearState.eIdle; // 回空闲 / back to idle
    ELSIF _fVbEst >= fVbLimitMm THEN // 越过寿命限值 / the life limit was passed
        _eState := E_DL_CncWearState.eChangeReq; // 迁换刀请求相 / migrate to the change request
    ELSIF _fVbEst < (_fAlarmMm - (fVbLimitMm * DL_CNC_HYST_BAND)) THEN // 回差带以下才降相（防抖）/ drop only below the hysteresis band
        IF _fVbEst >= fVbCompTrigMm THEN // 仍在补偿门限之上 / still above the trigger
            _eState := E_DL_CncWearState.eCompensate; // 降回补偿相 / drop back to compensating
        ELSE // 已回落到补偿门限之下 / fell below the trigger
            _eState := E_DL_CncWearState.eLearn; // 降回学习相 / drop back to learning
        END_IF
    END_IF
E_DL_CncWearState.eChangeReq: // 换刀请求相：锁存驻留，唯一解除为复位沿（段 3 已迁回空闲）
    IF NOT _bChangeLch THEN // 锁存已被复位沿清除 / the latch was cleared by the reset edge
        _eState := E_DL_CncWearState.eIdle; // 回空闲 / back to idle
    END_IF
ELSE // 非法相位兜底（R6、R128）/ the illegal phase fallback
    _eState := E_DL_CncWearState.eIdle; // 回安全态空闲 / back to the safe idle phase
    _iErrTmp := 2601; // 信息级非法相位码 / the info grade illegal phase code
END_CASE
IF _eState = E_DL_CncWearState.eChangeReq THEN _bChangeLch := TRUE; END_IF // 锁存单点置位（R187 两段式之一）/ single point latch set
// 段 10｜刀补增量闭环：状态量门控（R99），增量限幅 ±50 µm 每拍，累计上限 200 µm 单向
IF (_eState = E_DL_CncWearState.eCompensate) OR (_eState = E_DL_CncWearState.eAlarm) THEN // 仅补偿相与报警相出增量
    _fCompTgt := (_fVbEst - fVbCompTrigMm) * DL_CNC_UM_PER_MM; // 目标累计补偿量 [µm]，以补偿门限为零点 / the target accumulated compensation [um]
    IF _fCompTgt < 0.0 THEN _fCompTgt := 0.0; END_IF // 目标下限夹取（不回退已补量）/ the lower clamp, no retraction
    IF _fCompTgt > DL_CNC_ACC_UM THEN _fCompTgt := DL_CNC_ACC_UM; END_IF // 目标上限夹取 / the upper clamp
    _fStep := _fCompTgt - _fCompAcc; // 本拍应补增量 [µm] / the step required this scan [um]
    IF _fStep > DL_CNC_STEP_UM THEN _fStep := DL_CNC_STEP_UM; ELSIF _fStep < (0.0 - DL_CNC_STEP_UM) THEN _fStep := (0.0 - DL_CNC_STEP_UM); END_IF // 单拍双向限幅 / the two sided step limit
    _fCompAcc := _fCompAcc + _fStep; // 累计量单点写入（全库唯一写入点）/ the only write point of the accumulator
    IF _fCompAcc > DL_CNC_ACC_UM THEN _fCompAcc := DL_CNC_ACC_UM; END_IF // 累计上限硬钳 / the hard clamp of the accumulator
    IF _fCompAcc < 0.0 THEN _fCompAcc := 0.0; END_IF // 累计下限硬钳 / the hard clamp of the lower side
    fCompUm := _fStep; // 增量单点映射 / the single point mapping of the step
END_IF
// 段 11｜统一出口：输出单点映射，信息级码与有效性同源（R191 名实相符）
eState := _eState; // 相位单点映射 / the single point mapping of the phase
fVbEst := _fVbEst; // 估计单点映射 [mm] / the single point mapping of the estimate
fVbRaw := _fVbRaw; // 原值单点映射 [mm] / the single point mapping of the raw value
fCompAccUm := _fCompAcc; // 累计刀补单点映射 [µm] / the single point mapping of the accumulator
fPathM := _fPathM; // 路程单点映射 [m] / the single point mapping of the path
fKcRatio := _fRatio; // 比能比单点映射 [-] / the single point mapping of the ratio
xChangeReq := _bChangeLch; // 换刀请求回放锁存位 / replay the change request latch
xAlarm := (_eState = E_DL_CncWearState.eAlarm) OR (_eState = E_DL_CncWearState.eChangeReq); // 报警电平（含换刀请求相）/ the alarm level including the change request
iErrCode := _iErrTmp; // 信息级码单点映射（每拍重算，不锁存，R187）/ the info code mapping, recomputed every scan
xValid := _bValid AND (_iErrTmp = 0); // 有效性：判据全通过且无信息级异常 / valid when every gate passed and no info code is set
END_FUNCTION_BLOCK

(* ---- FB_DL_CoderRibbonLife.st ---- *)
(*
  FB_DL_CoderRibbonLife  —  打码机色带寿命双口径评估（次数口径 + 浓度口径取劣）/ Coder ribbon life, dual-criterion estimation
  分类 Category : DL_Device
  码位 Code     : 16#03_2_11
  版本 Version  : 1.0.0
  来源 Source   : t2-1-lgf-technology — IEC 61131-3 标准语义的道莅防御性实现
  溯源 Origin   : LGF 工艺类文档公开语义借鉴（耗材寿命双口径、浓度补偿），clean-room 实现，未复制源码行
  功能 Function : 1) 次数口径：已打次数 nPrintedCount 对额定 nRibbonRatingPrints 的余量 → fRemainCntPct；
                  2) 浓度口径：为达清晰度被迫把浓度指令抬升至 fDensityMinPct 之上的幅度，
                     超过 fDensityRiseMaxPct 即说明色带色粉已衰减 → fRemainDensPct（按抬升幅度线性折算）；
                  3) 两口径**取劣者**作为 fRemainPct 输出（任一口径到限即预警，不平均、不取优）；
                  4) bReplaceWarn 在 fRemainPct <= fWarnLevelPct 时置位（维护级告警，信息级 0121，不置 bError）；
                  5) bDensityCompSaturated 在浓度指令顶到 fDensityCeilPct（默认 100%）时置位（再无可调余量）。
  边界 Boundary : ① nRibbonRatingPrints = 0 判组态错 0211（次数口径的分母，R45 防除零）；
                      fDensityMinPct <= 0 / fDensityRiseMaxPct <= 0 / fWarnLevelPct 域外同判组态错；
                  ② fDensityCmdPct 越 0~100 时**钳制到域内**并置组态告警 0211（bError 置位，工艺参数错误
                     不允许静默通过）；钳制值参与后续全部换算，绝不用域外值做分母；
                  ③ nPrintedCount 为 UDINT，饱和到额定值**不回绕**（回绕会让色带寿命台账凭空复活）；
                     计数累加前做上限预判（R28-3：不写 TRUNC(x)+1，不靠事后比较）；
                  ④ 换带复位须 bRibbonReplaced 上升沿 **且** bReset 同时成立（解除式自证：两条件均可满足）；
                     只按 bRibbonReplaced 会丢掉操作员确认，只按 bReset 会把正常复位当成换带（台账污染）；
                  ⑤ bPrintPulse 用 R_TRIG 且**每主周期无条件刷新**（R182）；
                  ⑥ 浓度口径与次数口径的百分比均限幅到 [0, 100]（负余量不显示为负数，防 HMI 误解）。
  依赖 Depends  : 仅 Standard.library（TON / R_TRIG / ABS / MIN / MAX），零外部组件依赖
  同拍双窗配比  : 浓度告警去抖窗 tDensityDb 与心跳窗 DL_HEART_WINDOW 不同源；配比约束
                  tDensityDb <= DL_HEART_WINDOW，保证心跳窗内至少一次浓度结论更新（R100）

  码表 Error codes（本件格 03_2_11，子码步进 +0x10）:
    16#0003_0211 故障级：组态非法（额定次数 = 0 / 浓度基准 <= 0 / 抬升上限 <= 0 / 浓度指令越 0~100 已钳制）
    16#0003_0221 故障级：状态机落 ELSE 兜底（非法相位 ID）
    16#0003_0111 信息级：换带复位已执行（计数与口径全部归零，不置 bError）
    16#0003_0121 信息级：色带更换预警（维护级，fRemainPct <= fWarnLevelPct，不置 bError）
    16#0003_0131 信息级：浓度补偿已饱和（指令顶到上限，无再调余量，不置 bError）

  修订历史 Revision :
    2026-11-18  v1.0.0  R37 首版
*)

TYPE E_DL_RibbonState :
(
    eIdle  := 0,   // 空闲：未使能 / Idle, not enabled
    eRun   := 10,  // 运行：正常计数与评估 / Running, counting and evaluating
    eWarn  := 20,  // 预警：余量到限，仍可继续打印 / Warning, printing may continue
    eFault := 90   // 故障：组态非法锁定 / Fault, illegal configuration latched
);
END_TYPE

FUNCTION_BLOCK FB_DL_CoderRibbonLife
VAR_INPUT
    bEnable        : BOOL := FALSE;             // 总使能，FALSE 时不计次 / Master enable, low level stops counting
    bReset         : BOOL := FALSE;             // 复位，上升沿清故障锁存（与换带沿同时成立才清台账）/ Reset, clears the latch
    bRibbonReplaced : BOOL := FALSE;            // 换带完成信号（上升沿；须与 bReset 同拍才复位台账）/ Ribbon replaced, rising edge
    bPrintPulse    : BOOL := TRUE;              // 打印触发脉冲输入（上升沿计一次；R_TRIG 每拍无条件刷新）/ Print trigger, rising edge counts
    nRibbonRatingPrints : UDINT := 1000000;     // 色带额定打印次数 [次]，域 > 0 / Rated print count, domain above zero
    fDensityCmdPct : REAL := 60.0;              // 当前浓度指令 [%]，域 0~100 / Present density command [%]
    fDensityMinPct : REAL := 40.0;              // 浓度基准（新带所需浓度）[%]，域 > 0 / Density baseline of a new ribbon [%]
    fDensityRiseMaxPct : REAL := 40.0;          // 允许浓度抬升上限 [%]，域 > 0 / Permitted density rise [%]
    fDensityCeilPct : REAL := 100.0;            // 浓度上限（饱和判定点）[%]，域 > 基准 / Density ceiling for the saturation test [%]
    fWarnLevelPct  : REAL := 10.0;              // 更换预警余量门限 [%]，域 0~100 / Remaining-level warning threshold [%]
END_VAR
VAR_OUTPUT
    nPrintedCount  : UDINT;                     // 已打次数 [次]，饱和不超过额定值 / Printed count, saturated at the rating
    fRemainPct     : REAL;                      // 剩余寿命（双口径取劣）[%] / Remaining life, the worse of both criteria [%]
    fRemainCntPct  : REAL;                      // 次数口径余量 [%] / Remaining life by count [%]
    fRemainDensPct : REAL;                      // 浓度口径余量 [%] / Remaining life by density [%]
    bReplaceWarn   : BOOL;                      // 更换色带预警（维护级）/ Ribbon replacement warning
    bDensityCompSaturated : BOOL;               // 浓度补偿饱和 / Density compensation saturated
    bValid         : BOOL;                      // 判据可用标志 / Criteria usable
    bError         : BOOL;                      // 故障标志，派生自锁存 / Fault flag derived from the latch
    nErrId         : UDINT;                     // 事件码，0 = 无事件 / Event code, 0 = no event
    eStateOut      : E_DL_RibbonState;          // 状态出口，段尾单点映射 / State outlet, mapped at the tail
END_VAR
VAR
    tonHeart     : TON;                         // 周期心跳窗，自复位 / Periodic heartbeat window, self-resetting
    rtReset      : R_TRIG;                      // 复位上升沿 / Reset rising edge
    rtReplace    : R_TRIG;                      // 换带上升沿 / Replacement rising edge
    rtPrint      : R_TRIG;                      // 打印触发上升沿（每拍无条件刷新）/ Print rising edge, refreshed every scan
    _eState      : E_DL_RibbonState := E_DL_RibbonState.eIdle;  // 内部相位（CASE 唯一写入目标）/ Internal phase
    _uFault      : UDINT;                       // 故障码锁存 / Latched fault code
    _uInfo       : UDINT;                       // 信息码，每拍重算 / Information code, recomputed per scan
    _bFault      : BOOL;                        // 故障锁存位 / Latched fault bit
    _bCfgBad     : BOOL;                        // 组态非法聚合 / Configuration invalid aggregate
    _bDensClamped : BOOL;                       // 浓度指令被钳制 / The density command was clamped
    _nCountAcc   : UDINT;                       // 已打次数保持量 [次] / Held printed count
    _fDens       : REAL;                        // 生效浓度指令（钳制后）[%] / Effective density command [%]
    _fRisePct    : REAL;                        // 相对基准的浓度抬升 [%] / Density rise above the baseline [%]
    _fCntRemain  : REAL;                        // 次数口径余量 [%] / Remaining life by count [%]
    _fDensRemain : REAL;                        // 浓度口径余量 [%] / Remaining life by density [%]
    _fWorst      : REAL;                        // 双口径取劣结果 [%] / Worse criterion value [%]
    _bReplaceNow : BOOL;                        // 本拍更换预警判据成立 / Warning criterion present this scan
    _bHeartBrk   : BOOL := TRUE;                // 心跳窗断输入一拍 / One-scan heartbeat break
END_VAR
VAR CONSTANT
    DL_PCT_MAX    : REAL := 100.0;      // 百分比上限 [%] / Percentage ceiling
    DL_PCT_MIN    : REAL := 0.0;        // 百分比下限 [%] / Percentage floor
    DL_HEART_WINDOW : TIME := T#2S;     // 心跳观察窗 [ms]，自复位节拍 / Heartbeat window, self-resetting
    DL_COUNT_MAX  : UDINT := 16#FFFF_FFFE; // 次数硬上限（额定值异常放大时的兜底）[次] / Hard count ceiling
END_VAR

(* —— 段 0：定时器与边缘检测无条件周期刷新（R182：R_TRIG 必须在主体前部，不得置于 IF 内） —— *)
rtReset(CLK := bReset);                                          // 复位上升沿，每拍必调
rtReplace(CLK := bRibbonReplaced);                               // 换带上升沿，每拍必调
rtPrint(CLK := bPrintPulse);                                     // 打印上升沿，每拍必调（计数触发源）
tonHeart(IN := (NOT tonHeart.Q) AND (NOT _bHeartBrk), PT := DL_HEART_WINDOW);  // 心跳窗自复位
_bHeartBrk := FALSE;                                             // 断输入拍在调用后自清

(* —— 段 1：单拍量预清零（计数 / 口径保持量不入清单，R187①） —— *)
_uInfo       := 16#0000_0000;   // 信息码每拍重算
bError       := FALSE;          // 故障出口每拍重算，段 7 由锁存派生
bValid       := FALSE;          // 可用标志缺省 FALSE
bReplaceWarn := FALSE;          // 预警出口缺省 FALSE，段 8 单点置位
_bCfgBad     := FALSE;          // 组态非法预清零
_bDensClamped := FALSE;         // 浓度钳制标志预清零
_bReplaceNow := FALSE;          // 预警判据预清零

(* —— 段 2：复位沿与换带沿（台账复位为双条件，R28-1 解除式自证） —— *)
IF rtReset.Q THEN
    _bFault := FALSE;                // 复位沿清故障锁存位（台账不清，换带才清）
    _uFault := 16#0000_0000;         // 复位沿清锁存码
END_IF
IF rtReplace.Q AND rtReset.Q THEN
    _nCountAcc := 0;                 // 换带 + 复位同拍：已打次数归零
    _fCntRemain := DL_PCT_MAX;       // 次数口径余量回到 100 %
    _fDensRemain := DL_PCT_MAX;      // 浓度口径余量回到 100 %
    _uInfo := 16#0003_0111;          // 信息级：换带复位已执行
END_IF

(* —— 段 3：组态域闸（覆盖全部参与换算的引脚，R151） —— *)
IF nRibbonRatingPrints = 0 THEN
    _bCfgBad := TRUE;                // 额定次数为 0：次数口径分母非法（R45 防除零）
END_IF
IF (fDensityMinPct <> fDensityMinPct) OR (fDensityMinPct <= 0.0) OR (fDensityMinPct > DL_PCT_MAX) THEN
    _bCfgBad := TRUE;                // 浓度基准非法
END_IF
IF (fDensityRiseMaxPct <> fDensityRiseMaxPct) OR (fDensityRiseMaxPct <= 0.0) THEN
    _bCfgBad := TRUE;                // 允许抬升上限非法（浓度口径分母）
END_IF
IF (fDensityCeilPct <> fDensityCeilPct) OR (fDensityCeilPct <= fDensityMinPct) THEN
    _bCfgBad := TRUE;                // 浓度上限须严格大于基准（否则饱和判定无意义）
END_IF
IF (fWarnLevelPct <> fWarnLevelPct) OR (fWarnLevelPct < DL_PCT_MIN) OR (fWarnLevelPct > DL_PCT_MAX) THEN
    _bCfgBad := TRUE;                // 预警门限越 0~100 域
END_IF
_fDens := fDensityCmdPct;            // 生效浓度初值
IF (_fDens <> _fDens) THEN
    _bCfgBad := TRUE;                // 浓度指令非有限：无法解释
END_IF
IF _fDens > DL_PCT_MAX THEN
    _fDens := DL_PCT_MAX;            // 上钳制到域内（钳制值才参与换算）
    _bDensClamped := TRUE;           // 标记已钳制
END_IF
IF _fDens < DL_PCT_MIN THEN
    _fDens := DL_PCT_MIN;            // 下钳制
    _bDensClamped := TRUE;
END_IF
IF _bDensClamped THEN
    _bCfgBad := TRUE;                // 域外浓度：组态告警（工艺参数错误不得静默通过）
END_IF
IF _bCfgBad THEN
    _uFault := 16#0003_0211;         // 故障级：组态非法
    _bFault := TRUE;                 // 锁存位置位（复位沿可清）
    bError  := TRUE;                 // 故障标志置位（R45 配对）
    _eState := E_DL_RibbonState.eFault;  // 进故障相
END_IF

(* —— 段 4：次数累计（上限预判，饱和不回绕；禁用 TRUNC(x)+1 型写法） —— *)
IF rtPrint.Q AND bEnable AND (NOT _bFault) AND (NOT _bCfgBad) THEN
    IF _nCountAcc < nRibbonRatingPrints THEN
        IF _nCountAcc < DL_COUNT_MAX THEN
            _nCountAcc := _nCountAcc + 1;   // 计数 +1（双重上限：额定值与硬上限，均不回绕）
        END_IF
    END_IF
END_IF

(* —— 段 5：双口径余量计算（次数口径与浓度口径各自独立，取劣输出） —— *)
IF (NOT _bCfgBad) AND (nRibbonRatingPrints > 0) THEN
    _fCntRemain := (1.0 - (UDINT_TO_REAL(_nCountAcc) / UDINT_TO_REAL(nRibbonRatingPrints))) * DL_PCT_MAX;  // 次数口径余量 [%]
    IF _fCntRemain < DL_PCT_MIN THEN
        _fCntRemain := DL_PCT_MIN;                     // 下限保护（饱和计数时余量恰为 0）
    END_IF
    IF _fCntRemain > DL_PCT_MAX THEN
        _fCntRemain := DL_PCT_MAX;                     // 上限保护（计数小于额定时不超过 100）
    END_IF
    IF _fDens > fDensityMinPct THEN
        _fRisePct := (_fDens - fDensityMinPct) / fDensityMinPct * DL_PCT_MAX;   // 相对基准的抬升 [%]（分母已证 > 0）
    ELSE
        _fRisePct := 0.0;                              // 未抬升：无衰减指示
    END_IF
    IF _fRisePct >= fDensityRiseMaxPct THEN
        _fDensRemain := DL_PCT_MIN;                    // 抬升已达上限：浓度口径余量耗尽
    ELSE
        _fDensRemain := (1.0 - (_fRisePct / fDensityRiseMaxPct)) * DL_PCT_MAX;  // 线性折算余量 [%]（分母已证 > 0）
    END_IF
    IF _fDensRemain < DL_PCT_MIN THEN
        _fDensRemain := DL_PCT_MIN;                    // 下限保护
    END_IF
    IF _fDensRemain > DL_PCT_MAX THEN
        _fDensRemain := DL_PCT_MAX;                    // 上限保护
    END_IF
    _fWorst := MIN(_fCntRemain, _fDensRemain);         // 双口径取劣（任一到限即预警）
    _bReplaceNow := (_fWorst <= fWarnLevelPct);        // 预警判据
    IF _bReplaceNow AND (_eState <> E_DL_RibbonState.eFault) THEN
        _uInfo := 16#0003_0121;                        // 信息级：色带更换预警（维护级）
    END_IF
ELSE
    _fWorst := DL_PCT_MIN;                             // 组态非法：余量按最不利显示（不伪造 100 %）
END_IF

(* —— 段 6：相位机（只做迁移；出口在段 8） —— *)
CASE _eState OF

E_DL_RibbonState.eIdle:
    IF bEnable AND (NOT _bFault) AND (NOT _bCfgBad) THEN
        _eState := E_DL_RibbonState.eRun;              // 使能且组态合法：进运行相
    END_IF

E_DL_RibbonState.eRun:
    IF (NOT bEnable) THEN
        _eState := E_DL_RibbonState.eIdle;             // 失能：回空闲
    ELSIF _bReplaceNow THEN
        _eState := E_DL_RibbonState.eWarn;             // 余量到限：进预警相（仍允许打印）
    END_IF

E_DL_RibbonState.eWarn:
    IF (NOT bEnable) THEN
        _eState := E_DL_RibbonState.eIdle;             // 失能：回空闲
    ELSIF (NOT _bReplaceNow) AND (rtReplace.Q AND rtReset.Q) THEN
        _eState := E_DL_RibbonState.eRun;              // 换带复位完成：回运行相
    END_IF

E_DL_RibbonState.eFault:
    IF (NOT _bFault) AND (NOT _bCfgBad) AND bEnable THEN
        _eState := E_DL_RibbonState.eRun;              // 锁存已清且组态合法：回运行相
    END_IF

ELSE
    _uFault := 16#0003_0221;                           // 故障级：相位 ID 越界（枚举兜底）
    _bFault := TRUE;                                   // 锁存
    bError  := TRUE;                                   // 故障标志置位（R45 配对）
    _eState := E_DL_RibbonState.eFault;                // 强制回故障相
END_CASE

(* —— 段 7：故障码优先级链（每个 bError 置位源在此均有码，R45 配对） —— *)
IF _bCfgBad THEN
    _uFault := 16#0003_0211;                           // 组态非法优先上报
    _bFault := TRUE;
    bError  := TRUE;
END_IF

(* —— 段 8：出口单点映射（名实同源；锁存码回放，禁同拍抹除） —— *)
nPrintedCount  := _nCountAcc;                          // 已打次数出口（饱和）
fRemainCntPct  := _fCntRemain;                         // 次数口径余量出口
fRemainDensPct := _fDensRemain;                        // 浓度口径余量出口
fRemainPct     := _fWorst;                             // 双口径取劣余量出口
bReplaceWarn   := (_eState = E_DL_RibbonState.eWarn);  // 预警出口（状态派生，与 eWarn 相严格同源）
bDensityCompSaturated := (_fDens >= fDensityCeilPct) AND (NOT _bCfgBad);  // 浓度补偿饱和：指令顶到上限
IF bDensityCompSaturated THEN
    _uInfo := 16#0003_0131;                            // 信息级：浓度补偿已饱和（无再调余量）
END_IF
eStateOut := _eState;                                  // 状态出口
IF _bFault THEN
    nErrId := _uFault;                                 // 故障锁存码回放（不在故障相按当下输入重推）
    bError := TRUE;                                    // 故障出口派生自锁存
ELSE
    nErrId := _uInfo;                                  // 信息码
END_IF
bValid := bEnable AND (NOT _bFault) AND (NOT _bCfgBad);  // 判据可用

END_FUNCTION_BLOCK

(* ---- FB_DL_CoilCarIndexSeq.st ---- *)
(*
  Name: FB_DL_CoilCarIndexSeq
  Category: DL_Device
  Version: 1.0.0
  Round: R89 / 2026-11-25
  开源溯源：clean-room 自研（族 板带剪切分条卷取，ST 开源生态实测 0 命中，无外部代码引入）
  功能：钢卷小车行走定位顺控（快进→慢进→精定位→落卷→返回），五相各自独立超时 TON。
  边界条件：① 位置与公差入参全部过非有限闸；配置越域即故障（101）；
            ② 快进/慢进/精定位/返回四相各用独立 TON，落卷为确定性时窗 DL_CCS_DROP，禁跨相共用（R100）；
            ③ 位置判据假设小车前进方向为位置数值增大（fPosSlowMm < fPosTargetMm），越序即组态非法；
            ④ 故障解除唯一路径：故障相内 xStart 释放（R152），清锁存回 eIdle。
  状态机：eIdle / eFast / eSlow / eFine / eDrop / eReturn / eDone / eFault（CASE 含 ELSE 兜底）。
*)
TYPE E_DL_CcsPhase :
(
    eIdle   := 0,       (* 待机：等启动沿 / Idle, waiting for start edge *)
    eFast   := 10,      (* 快进相：走到减速点 / Fast travel to slow-down point *)
    eSlow   := 20,      (* 慢进相：走到精定位带 / Slow travel to fine band *)
    eFine   := 30,      (* 精定位相：进入公差带 / Fine positioning into tolerance *)
    eDrop    := 40,     (* 落卷相：确定性落卷时窗 / Coil drop, fixed window *)
    eReturn := 50,      (* 返回相：回到原点位 / Return to home position *)
    eDone    := 60,     (* 完成相：保持至启动释放 / Done, holds until start released *)
    eFault  := 90       (* 故障相：锁存待释放 / Fault latched, awaiting release *)
);
END_TYPE

FUNCTION_BLOCK FB_DL_CoilCarIndexSeq
VAR_INPUT
    xStart : BOOL;          (* 启动命令（上升沿起序） [-] Start command, rising edge *)
    fPosActMm : REAL;       (* 小车位置实测 [mm] Car position actual [mm] *)
    fPosSlowMm : REAL;      (* 减速（慢进）点位置 [mm] Slow-down point [mm] *)
    fPosTargetMm : REAL;    (* 精定位目标位置 [mm] Fine positioning target [mm] *)
    fTolMm : REAL;          (* 精定位公差 [mm] Fine positioning tolerance [mm] *)
    tTimeoutS : TIME;       (* 单相超时窗 [ms] Phase timeout window [ms] *)
END_VAR
VAR_OUTPUT
    eState : E_DL_CcsPhase; (* 当前相 [-] Present phase *)
    xDone : BOOL;           (* 完成单拍脉冲 [-] One-scan done pulse *)
    xFault : BOOL;          (* 故障锁存标志 [-] Fault latched *)
    nErrCode : INT;         (* 故障码 0/101 组态/102~105 超时/106 非法相 [-] Error code *)
END_VAR
VAR
    _ePhase : E_DL_CcsPhase := E_DL_CcsPhase.eIdle;  (* 内部相（CASE 唯一写入目标） [-] Internal phase *)
    _bDone : BOOL := FALSE;         (* 单拍完成标志（段 1 预清） [-] One-scan done flag *)
    _bFaultLatch : BOOL := FALSE;   (* 故障锁存位 [-] Fault latch *)
    _bReqFault : BOOL := FALSE;     (* 单拍故障请求（段 1 预清） [-] Fault request *)
    _bCfgBad : BOOL := FALSE;       (* 组态非法当拍量 [-] Configuration bad *)
    _nErr : INT := 0;               (* 故障码锁存 [-] Latched error code *)
    _nReqErr : INT := 0;            (* 当拍请求码 [-] Requested error code *)
    _fErrMm : REAL := 0.0;          (* 距目标偏差绝对量 [mm] Absolute deviation to target [mm] *)
    tonFast : TON;                  (* 快进超时（段 0 无条件调用） / Fast travel timeout *)
    tonSlow : TON;                  (* 慢进超时（段 0 无条件调用） / Slow travel timeout *)
    tonFine : TON;                  (* 精定位超时（段 0 无条件调用） / Fine positioning timeout *)
    tonDrop : TON;                  (* 落卷时窗（确定性时窗） / Coil drop window *)
    tonReturn : TON;                (* 返回超时（段 0 无条件调用） / Return timeout *)
    rtStart : R_TRIG;               (* 启动沿（段 0 无条件调用） / Start edge *)
END_VAR
VAR CONSTANT
    DL_CCS_SLOW_BAND : REAL := 5.0;         (* 精定位带半宽（取 5 倍公差不劣于公差） [mm] Fine band half-width [mm] *)
    DL_CCS_HOME_MM : REAL := 10.0;          (* 原点位判定门限 [mm] Home position threshold [mm] *)
    DL_CCS_DROP : TIME := T#800MS;          (* 落卷动作时窗（确定性） [ms] Coil drop window [ms] *)
END_VAR
(* —— 段 0：沿与五 TON 无条件周期刷新（R7），IN 仅由相位派生 —— *)
rtStart(CLK := xStart);                                             (* 启动沿 / Start edge *)
tonFast(IN := (_ePhase = E_DL_CcsPhase.eFast), PT := tTimeoutS);    (* 快进超时 / Fast timeout *)
tonSlow(IN := (_ePhase = E_DL_CcsPhase.eSlow), PT := tTimeoutS);    (* 慢进超时 / Slow timeout *)
tonFine(IN := (_ePhase = E_DL_CcsPhase.eFine), PT := tTimeoutS);    (* 精定位超时 / Fine timeout *)
tonDrop(IN := (_ePhase = E_DL_CcsPhase.eDrop), PT := DL_CCS_DROP);  (* 落卷时窗 / Drop window *)
tonReturn(IN := (_ePhase = E_DL_CcsPhase.eReturn), PT := tTimeoutS);(* 返回超时 / Return timeout *)
(* 非有限闸（NaN 自反 + Inf 差值自减）+ 组态域闸：位置与公差全枚举（R272） *)
_bCfgBad := (fPosActMm <> fPosActMm) OR ((fPosActMm - fPosActMm) <> 0.0)
         OR (fPosSlowMm <> fPosSlowMm) OR ((fPosSlowMm - fPosSlowMm) <> 0.0)
         OR (fPosTargetMm <> fPosTargetMm) OR ((fPosTargetMm - fPosTargetMm) <> 0.0)
         OR (fTolMm <> fTolMm) OR ((fTolMm - fTolMm) <> 0.0)
         OR (fTolMm < 0.1) OR (fTolMm > 20.0)
         OR (fPosSlowMm >= fPosTargetMm) OR (fPosTargetMm > 30000.0) OR (tTimeoutS <= T#0S);
(* 偏差绝对量：容差比较一律用差值，禁浮点判等 *)
_fErrMm := ABS(fPosActMm - fPosTargetMm);
(* —— 段 1：单拍量预清零 —— *)
_bDone := FALSE;
_bReqFault := FALSE;
_nReqErr := 0;
IF _bCfgBad THEN
    _bReqFault := TRUE; _nReqErr := 101;        (* 组态非法 / Configuration bad *)
END_IF
(* —— 段 2：故障锁存解除（唯一路径 = 故障相内 xStart 释放，R152） —— *)
IF _bFaultLatch AND (NOT xStart) THEN
    _bFaultLatch := FALSE;                      (* 清锁存 / Clear latch *)
    _nErr := 0;                                 (* 清码 / Clear code *)
    _ePhase := E_DL_CcsPhase.eIdle;             (* 迁回待机 / Back to idle *)
END_IF
(* —— 段 3：主状态机（ENUM + CASE，ELSE 兜底） —— *)
CASE _ePhase OF
E_DL_CcsPhase.eIdle:
    IF rtStart.Q AND (NOT _bFaultLatch) THEN
        _ePhase := E_DL_CcsPhase.eFast;         (* 起序 → 快进 / Start to fast travel *)
    END_IF
E_DL_CcsPhase.eFast:
    IF fPosActMm >= fPosSlowMm THEN
        _ePhase := E_DL_CcsPhase.eSlow;         (* 到减速点 → 慢进 / Reached slow-down point *)
    ELSIF tonFast.Q THEN
        _bReqFault := TRUE; _nReqErr := 102;    (* 快进超时 / Fast travel timeout *)
    END_IF
E_DL_CcsPhase.eSlow:
    IF _fErrMm <= DL_CCS_SLOW_BAND THEN
        _ePhase := E_DL_CcsPhase.eFine;         (* 进精定位带 → 精定位 / Enter fine band *)
    ELSIF tonSlow.Q THEN
        _bReqFault := TRUE; _nReqErr := 103;    (* 慢进超时 / Slow travel timeout *)
    END_IF
E_DL_CcsPhase.eFine:
    IF _fErrMm <= fTolMm THEN
        _ePhase := E_DL_CcsPhase.eDrop;         (* 进公差带 → 落卷 / In tolerance, drop *)
    ELSIF tonFine.Q THEN
        _bReqFault := TRUE; _nReqErr := 104;    (* 精定位超时 / Fine positioning timeout *)
    END_IF
E_DL_CcsPhase.eDrop:
    IF tonDrop.Q THEN
        _ePhase := E_DL_CcsPhase.eReturn;       (* 落卷时窗到 → 返回 / Drop done, return *)
    END_IF
E_DL_CcsPhase.eReturn:
    IF fPosActMm <= DL_CCS_HOME_MM THEN
        _bDone := TRUE;                         (* 单拍完成（段 1 预清） / One-scan done *)
        _ePhase := E_DL_CcsPhase.eDone;         (* → 完成相 / To done *)
    ELSIF tonReturn.Q THEN
        _bReqFault := TRUE; _nReqErr := 105;    (* 返回超时 / Return timeout *)
    END_IF
E_DL_CcsPhase.eDone:
    IF NOT xStart THEN
        _ePhase := E_DL_CcsPhase.eIdle;         (* 启动释放 → 待机 / Start released, idle *)
    END_IF
E_DL_CcsPhase.eFault:
    _fErrMm := ABS(fPosActMm - fPosTargetMm);   (* 故障相驻留：仅刷新偏差量供追溯，不迁相 *)
ELSE
    _bReqFault := TRUE;                         (* 非法相兜底 / Illegal phase fallback *)
    _nReqErr := 106;
END_CASE
(* —— 段 4：故障请求统一落地（唯一锁存点 + 同步迁相，R187/R252） —— *)
IF _bReqFault AND (NOT _bFaultLatch) THEN
    _bFaultLatch := TRUE;                       (* 锁存 / Latch *)
    _nErr := _nReqErr;                          (* 码锁存回放 / Latched code *)
    _ePhase := E_DL_CcsPhase.eFault;            (* 同步迁相 / Migrate to fault *)
END_IF
(* —— 段 5：统一出口（各出口单点赋值） —— *)
eState := _ePhase;
xDone := _bDone;
xFault := _bFaultLatch;
nErrCode := _nErr;
END_FUNCTION_BLOCK

(* ---- FB_DL_CoilFreezeStat.st ---- *)
// =====================================================================
// FB_DL_CoilFreezeStat.st
// 盘管防冻统计判据（只判不控：低温累计 + 温降速率，预警/报警锁存）
// Coil freeze statistics FB (detect only)
// 码位: 16#0003_03CA ~ 16#0003_03CE (本件独占 5 槽)
// 修改记录: R29 初版 (按 DISPATCH_R29 序 9)
// =====================================================================
FUNCTION_BLOCK FB_DL_CoilFreezeStat
VAR_INPUT
    bEnable        : BOOL  := FALSE;   // 使能 / Enable
    bReset         : BOOL  := FALSE;   // 复位锁存 / Reset
    bTempValid     : BOOL  := FALSE;   // 温度有效 / Temp valid
    fCoilTemp_C    : REAL  := 12.0;    // 盘管温度 -40~80 ℃ / Coil temperature [degC]
    fFreezeLimit_C : REAL  := 2.0;     // 冻结判定限 -10~10 ℃ / Freeze limit [degC]
    fRateAlarm_Cmin : REAL := 1.0;     // 温降速率报警 0.1~20 K/min / Cooling rate alarm [K/min]
    tAccumWarn     : TIME  := T#5M;    // 累计预警 T#10S~T#2H / Accumulate warn [s]
    tAccumAlarm    : TIME  := T#10M;   // 累计报警 T#10S~T#8H / Accumulate alarm [s]
    fDecayFactor   : REAL  := 0.5;     // 回暖衰减系数 0~1 / Decay factor [-]
    bFanRun        : BOOL  := FALSE;   // 风机运行 / Fan running
    tCycle         : TIME  := T#1S;    // 周期 T#100MS~T#10S / Cycle [s]
END_VAR
VAR_OUTPUT
    tColdAccum     : TIME;             // 低温累计时长 / Cold accumulate [s]
    fRate_Cmin     : REAL;             // 温降速率 K/min / Cooling rate [K/min]
    bWarn          : BOOL;             // 预警 / Warning
    bAlarm         : BOOL;             // 报警（锁存）/ Alarm latched
    eErr           : UDINT;            // 错误码 / Error code
END_VAR
VAR
    fTempPrev      : REAL  := 12.0;    // 上拍温度快照 / Previous temperature snapshot [degC]
    fTempAcc       : REAL  := 0.0;     // 累计秒值（内部实数实现）/ Accumulated seconds, internal [s]
    tWarnS         : REAL;             // 预警阈值秒 / Warn threshold seconds [s]
    tAlarmS        : REAL;             // 报警阈值秒 / Alarm threshold seconds [s]
    tCycleS        : REAL;             // 周期秒值（钳 ≥0.1）/ Cycle seconds, clamped [s]
    fDelta         : REAL;             // 温度差 / Temperature delta [K]
    fRateRaw       : REAL;             // 原始速率 K/min / Raw rate [K/min]
    fRateMaxLim    : REAL;             // 速率显示上限 / Rate display limit [K/min]
    bRateTrip      : BOOL;             // 速率越限 / Rate trip flag
    tAccumUpperS   : REAL;             // 累计上界 = 2×报警阈值 / Accum upper bound [s]
    bDecayOK       : BOOL;             // 衰减可执行标记 / Decay allowed flag
    xFirstScan     : BOOL  := TRUE;    // 首扫标记 / First-scan flag
END_VAR

// ---------------------------------------------------------------------
// 代码位表（本件独占，勿复用）:
//   16#0003_03CA 信息 统计正常（未越限）
//   16#0003_03CB 故障 温度非有限 / tCycle 非法
//   16#0003_03CC 故障 tAccumAlarm ≤ tAccumWarn / fDecayFactor < 0 / fDecayFactor > 1（组态错）
//   16#0003_03CD 信息 bTempValid=FALSE → 累计冻结（不增不减）
//   16#0003_03CE 故障 tColdAccum ≥ tAccumAlarm 或 fRate_Cmin ≥ fRateAlarm_Cmin → bAlarm=TRUE 锁存
// ---------------------------------------------------------------------

// ---- 周期与阈值转秒 / Cycle and thresholds to seconds ----
tCycleS  := TIME_TO_REAL(tCycle) / 1000.0;      // 周期秒值 / Cycle seconds [s]
tWarnS   := TIME_TO_REAL(tAccumWarn) / 1000.0;  // 预警阈值秒 / Warn threshold [s]
tAlarmS  := TIME_TO_REAL(tAccumAlarm) / 1000.0; // 报警阈值秒 / Alarm threshold [s]
IF tCycleS < 0.1 THEN
    tCycleS := 0.1;             // 钳 ≥0.1 s 防差分噪声放大 / Clamp 0.1 s min
END_IF

// ---- 非有限与周期合法性闸 / Finite and cycle validity gate ----
IF (tCycle = T#0MS) OR (tCycleS > 10.0)
   OR (fCoilTemp_C <> fCoilTemp_C) OR (ABS(fCoilTemp_C) >= 1.0E12) THEN
    eErr := 16#0003_03CB;       // 故障码 / Fault code
    RETURN;                     // 累计与报警保持 / Accum and alarm hold
END_IF

// ---- 组态错闸 / Configuration fault gate ----
IF (tAccumAlarm <= tAccumWarn) OR (fDecayFactor < 0.0) OR (fDecayFactor > 1.0)
   OR (fRateAlarm_Cmin <= 0.0) THEN
    eErr := 16#0003_03CC;       // 故障码 / Fault code
    RETURN;                     // 本拍结束 / End of cycle
END_IF

// ---- 累计上界 / Accum upper bound ----
tAccumUpperS := 2.0 * tAlarmS;  // 上界 = 2×报警阈值 / Upper bound 2x alarm

// ---- 首扫初始化（R16 首扫纪律）/ First-scan initialization ----
IF xFirstScan THEN
    fTempPrev := fCoilTemp_C;   // 快照对齐当前 / Snapshot align
    xFirstScan := FALSE;        // 清标记 / Clear flag
END_IF

// ---- 使能撤销：累计与报警保持，速率清零 / Disable: hold accum, zero rate ----
IF NOT bEnable THEN
    fRate_Cmin := 0.0;          // 速率清零 / Rate zero
    bWarn := FALSE;             // 预警复位 / Warn reset
    eErr := 16#0003_03CA;       // 信息级：空闲正常 / Info: idle normal
    RETURN;                     // 累计与报警锁存保持 / Accum and latch hold
END_IF

// ---- 温度传感器无效 → 冻结累计（不增不减）+ 信息级 / Temp invalid: freeze accum ----
IF NOT bTempValid THEN
    eErr := 16#0003_03CD;       // 信息级：累计冻结 / Info: accum frozen
    fTempPrev := fCoilTemp_C;   // 快照对齐防恢复瞬跳 / Align snapshot to avoid spike
    RETURN;                     // 累计与报警保持 / Accum and alarm hold
END_IF

// ---- 温降速率（一阶差分）/ Cooling rate (first-order difference) ----
fDelta := fCoilTemp_C - fTempPrev;          // 温度差 / Temperature delta [K]
fRateRaw := -fDelta / (tCycleS / 60.0);     // 降温为正，K/min / Positive when cooling [K/min]
IF fRateRaw > 1.0E12 THEN
    fRateRaw := 1.0E12;         // 速率显示上限防溢出 / Rate display clamp
END_IF
fRate_Cmin := fRateRaw;         // 输出速率 / Output rate

// ---- 速率越限判（即使累计未到）/ Rate trip check (even if accum low) ----
bRateTrip := (fRateRaw >= fRateAlarm_Cmin);     // 越限标志 / Trip flag

// ---- 累计逻辑：低温累计，回暖衰减 / Accumulation: cold add, warm decay ----
bDecayOK := FALSE;              // 衰减标记复位 / Reset flag
IF fCoilTemp_C < fFreezeLimit_C THEN
    // 低温：累计递增 / Cold: accumulate
    fTempAcc := fTempAcc + tCycleS;     // 累加 / Add cycle
    IF fTempAcc > tAccumUpperS THEN
        fTempAcc := tAccumUpperS;       // 钳上界防溢出 / Clamp upper bound
    END_IF
ELSE
    // 回暖且风机运行：按衰减系数递减（不得低于 0）/ Warm + fan: decay, floor 0
    IF bFanRun AND (fTempAcc > 0.0) THEN
        fTempAcc := fTempAcc - fDecayFactor * tCycleS;  // 衰减 / Decay
        IF fTempAcc < 0.0 THEN
            fTempAcc := 0.0;    // 下限 0 / Floor 0
        END_IF
        bDecayOK := TRUE;       // 衰减已执行 / Decay executed
    END_IF
END_IF
tColdAccum := REAL_TO_TIME(fTempAcc * 1000.0);  // 输出累计时长 / Output accumulate

// ---- 报警锁存 / Alarm latch ----
IF bRateTrip OR (fTempAcc >= tAlarmS) THEN
    bAlarm := TRUE;             // 锁存 / Latch
END_IF

// ---- 锁存解除式（可达性自证：三条件齐才解除，R28）/ Release path: all three conditions ----
IF bAlarm AND bReset
   AND (fCoilTemp_C > fFreezeLimit_C + 2.0)
   AND (fRate_Cmin < 0.0) THEN
    bAlarm := FALSE;            // 解除报警锁存 / Release alarm latch
    fTempAcc := 0.0;            // 累计清零 / Accum cleared
    tColdAccum := T#0MS;        // 输出同步清零 / Output synced
END_IF

// ---- 预警与错误码（故障级优先，锁存回放不重推断）/ Warn and code, fault replay first ----
IF bAlarm THEN
    bWarn := TRUE;              // 报警含预警 / Alarm implies warn
    eErr  := 16#0003_03CE;      // 故障码回放 / Fault code replay
ELSE
    bWarn := (fTempAcc >= tWarnS);  // 累计预警判 / Accum warn verdict
    IF bWarn THEN
        eErr := 16#0003_03CA;   // 信息级：预警期统计正常口径 / Info: warn period
    ELSE
        eErr := 16#0003_03CA;   // 信息级：统计正常 / Info: normal
    END_IF
END_IF

// ---- 上拍快照更新 / Previous snapshot update ----
fTempPrev := fCoilTemp_C;       // 快照 / Snapshot

END_FUNCTION_BLOCK

(* ---- FB_DL_CoilFrostWindow.st ---- *)
//==============================================================================
// 功能块：FB_DL_CoilFrostWindow ｜ 中文名称：盘管结霜窗口判定与除霜请求
// 所属子库：DL_Device ｜ 版本：v1.0.0 ｜ 兼容：CODESYS V3.5+ / TwinCAT 3 / 汇川 InoProShop
// 功能描述：结霜双判据窗——盘管表面温度同时满足「冻结判据」（表面温度
//           <= 结霜阈值）与「露点判据」（表面温度 <= 露点 - 裕度，有凝
//           才有霜）持续 tFrostDwell → 结霜窗确认，锁存除霜请求；除霜
//           完成判据 = 表面温度 > 结霜阈值 + 回差 fThawHystK（退出回差，
//           阈值附近抖动防频动，R23 教训同理）。露点由 Magnus-Tetens
//           内联解算（Device 不得调用 DL_Algo，见依赖纪律）。
// 开源溯源 (Origin)：道莅原创实现（参考换热盘管结霜判据与除霜控制工程惯例 分类与参数域）
// 单位表：温度[摄氏度] / 露点[摄氏度] / 裕度与回差[开] / 时间[ms]
// 错误码表：16#0003_018A 信息级（结霜窗确认、除霜请求锁存建立，不置
//           bError）/ 16#0003_018B 信息级（除霜完成回差退出，请求解除，
//           不置 bError）/ 16#0003_0360 故障级（组态非法：阈值/裕度/
//           回差域、时间窗 <= 0 或任一输入非有限，置 bError）/
//           16#0003_0361 故障级（传感器交叉校验失败：解算露点 > 干球
//           + 1 开，物理不可能，判湿度/温度通道异常，安全侧锁存除霜
//           请求，置 bError——该场景不可由 0360 的组态类判据观测，
//           属运行数据独立域）/ 16#0003_0362 故障级兜底（状态机落 ELSE，
//           置 bError）
// 状态机：E_DL_CoilFrostState（五态：eIdle=0 / eMonitor=10 / eFrost=20 /
//           eDefrost=30 / eFault=99），CASE 含 ELSE 兜底，ELSE 置 0362
// 边界行为：① 组态非法 → 故障态锁存，bReset 复位；② 湿度域外钳
//           1~100 照算（Magnus 对数域下限保证）；③ 驻留窗未满判据消失
//           → 自动回监视态（防瞬时低温误锁存）；④ 除霜请求锁存后仅
//           回差退出或 bReset 解除；⑤ 未使能输出冻结零并 bValid :=
//           FALSE（除霜请求不在未使能态保持——使能即监视语义）；⑥
//           安全侧 = 交叉校验失败时锁存除霜请求（宁多除一次，不漏霜）。
// 依赖纪律：Device 不得调用 DL_Algo——Magnus-Tetens 露点解算在本件内联
//           实现，常量口径（17.62/243.12/611.2）与 FC_DL_AirDensity
//           族一致性由本件头注释承担验证责任，改动任一侧须复核另一侧。
// 修订历史：v1.0.0 2026-11-17 首版（R24 派单 · ROADMAP P1 §727）
//==============================================================================

(*------------------------------------------------------------------------------
 * 枚举: E_DL_CoilFrostState（归属本功能块，同文件发布，全库唯一定义）
 * 含义: 结霜监视相位，每个成员在 CASE 中有且仅有一个标签。
 *-----------------------------------------------------------------------------*)
TYPE E_DL_CoilFrostState :
(
    eIdle    := 0,   // 空闲：未使能 / Idle, not enabled
    eMonitor := 10,  // 监视：判据计窗中 / Monitor, criteria window counting
    eFrost   := 20,  // 霜窗：双判据持续驻留已确认 / Frost, dual-criteria dwell confirmed
    eDefrost := 30,  // 除霜：请求锁存保持，等回差退出 / Defrost, request latched, awaiting the hysteresis exit
    eFault   := 99   // 故障：组态非法/交叉校验/非法状态 / Fault, config, cross-check or illegal state
);
END_TYPE

FUNCTION_BLOCK FB_DL_CoilFrostWindow
VAR_INPUT
    bEnable         : BOOL;                 // 监视使能 [—] / Monitoring enable
    bReset          : BOOL;                 // 故障复位 [—]，上升沿清锁存 / Fault reset, rising edge clears latches
    fAirTempC       : LREAL;                // 空气干球温度 [摄氏度] / Air dry-bulb temperature [degC]
    fRhPct          : LREAL;                // 空气相对湿度 [百分数]，域外钳 1..100 照算 / Air relative humidity [percent], clamped 1..100
    fCoilSurfTempC  : LREAL;                // 盘管表面温度 [摄氏度] / Coil surface temperature [degC]
    fFrostThreshC   : LREAL := 0.0;         // 结霜阈值 [摄氏度]，表面低于此判冻结 / Frost threshold [degC], freezing below
    fDpMarginK      : LREAL := 1.0;         // 露点裕度 [开]，表面低于露点减此值判凝露 / Dew-point margin [K]
    fThawHystK      : LREAL := 2.0;         // 除霜退出回差 [开]，须 > 0 且 < 裕度 + 10 / Thaw hysteresis [K], exit band width
    tFrostDwell     : TIME  := T#60S;       // 双判据驻留窗 [ms]，须 > 0 / Dual-criteria dwell window [ms]
END_VAR
VAR_OUTPUT
    fDewPointC      : LREAL;                // 解算露点 [摄氏度]（诊断出口） / Solved dew point [degC], diagnostics outlet
    bFrostWindow    : BOOL;                 // 结霜窗判定中 [—]（霜窗态电平） / Frost-window active level
    bDefrostReq     : BOOL;                 // 除霜请求 [—]（锁存保持） / Defrost request, latched
    eState          : E_DL_CoilFrostState;  // 相位出口 [—] / Phase outlet
    eErr            : UDINT;                // 错误码，0 = 无错，码位 16#0003_018A 起信息级、16#0003_0360 起故障级（分带见错误码表） / Error code, 0 = no error, band info/fault per the code table
    bError          : BOOL;                 // 故障级标志，仅故障级错误置位 / Fault-class flag, set only on fault-level codes
    bValid          : BOOL;                 // 输出可用标志 / Outputs usable flag
END_VAR
VAR
    fbDwell     : TON;                      // 双判据驻留计时（每拍无条件刷新）[ms] / Dwell timer, refreshed unconditionally
    _eState     : E_DL_CoilFrostState := E_DL_CoilFrostState.eIdle; // 当前相位 / Current phase
    _bCfgBad    : BOOL;                     // 组态非法锁存 / Illegal config latch
    _bCrossBad  : BOOL;                     // 交叉校验失败锁存 / Cross-check fault latch
    _bInfoFrost : BOOL;                     // 霜窗信息当拍标志 / Frost-window info flag of this scan
    _bInfoDone  : BOOL;                     // 除霜完成信息当拍标志 / Defrost-done info flag of this scan
    _bDefrostL  : BOOL;                     // 除霜请求锁存 / Defrost request latch
    _fRhUse     : LREAL;                    // 生效湿度（已钳位）[百分数] / Effective humidity, clamped
    _fGamma     : LREAL;                    // 露点解算中间量 ln(RH/100) [无量纲] / Dew-point intermediate ln(RH/100)
    _fDpCalc    : LREAL;                    // 解算露点 [摄氏度] / Solved dew point [degC]
    _bIllegal   : BOOL;                     // 非法状态标志 / Illegal state flag
    _bInit      : BOOL := FALSE;            // 首扫标志，初值 FALSE 取非判定 / First-scan flag, tested negated
END_VAR
VAR CONSTANT
    DL_CFW_MAGNUS_A : LREAL := 17.62;       // Magnus 系数 A [无量纲]，与 FC_DL_AirDensity 同口径 / Magnus coefficient A, aligned with FC_DL_AirDensity
    DL_CFW_MAGNUS_B : LREAL := 243.12;      // Magnus 系数 B [摄氏度]，同口径 / Magnus coefficient B, aligned
    DL_CFW_INF      : LREAL := 1.7976931348623157E308; // LREAL 幅值上限 / LREAL magnitude ceiling
    DL_CFW_EPS      : LREAL := 1.0E-6;      // 浮点判零容差 [混合] / Float zero tolerance
    DL_CFW_RH_MIN   : LREAL := 1.0;         // 湿度钳位下限 [百分数]（对数域保证） / Humidity clamp floor [percent]
    DL_CFW_RH_MAX   : LREAL := 100.0;       // 湿度钳位上限 [百分数] / Humidity clamp ceiling [percent]
    DL_CFW_CROSS_K  : LREAL := 1.0;         // 交叉校验容差 [开]（露点 > 干球 + 此值判异常） / Cross-check tolerance [K]
    DL_CFW_ZERO     : LREAL := 0.0;         // 零值常量，避免裸字面量 [混合] / Zero constant, avoids a bare literal
END_VAR

(*------------------------------------------------------------------------------
 * 段 1｜每拍预置：输出安全侧清零，单拍标志预清零
 *      Outputs cleared fail-safe first, one-shot flags pre-cleared
 *-----------------------------------------------------------------------------*)
fDewPointC   := DL_CFW_ZERO;             // 露点出口先清 / Dew point cleared first
bFrostWindow := FALSE;                   // 霜窗电平先清 / Frost level cleared first
eErr   := 16#0000_0000;                  // 错误码每拍重算 / Error code recomputed
bError := FALSE;                         // 故障标志每拍重算 / Fault flag recomputed
bValid := FALSE;                         // 可用标志每拍重算 / Usable flag recomputed
_bInfoFrost := FALSE;                    // 霜窗信息预清零 / Frost info pre-cleared
_bInfoDone  := FALSE;                    // 完成信息预清零 / Done info pre-cleared
_bIllegal   := FALSE;                    // 非法状态预清零 / Illegal flag pre-cleared

(*------------------------------------------------------------------------------
 * 段 2｜首扫初始化
 *      First-scan initialisation
 *-----------------------------------------------------------------------------*)
IF NOT _bInit THEN
    _eState    := E_DL_CoilFrostState.eIdle; // 相位空闲起步 / Phase starts idle
    _bCfgBad   := FALSE;                 // 组态锁存清零 / Config latch cleared
    _bCrossBad := FALSE;                 // 交叉锁存清零 / Cross latch cleared
    _bDefrostL := FALSE;                 // 请求锁存清零 / Request latch cleared
    _bInit     := TRUE;                  // 首扫只做一次 / The first scan runs once
END_IF

(*------------------------------------------------------------------------------
 * 段 3｜组态防御闸：非有限（R79）+ 阈值/裕度/回差/时间窗域
 *      Configuration defense gates
 *-----------------------------------------------------------------------------*)
IF (fAirTempC <> fAirTempC) OR (ABS(fAirTempC) > DL_CFW_INF)
   OR (fRhPct <> fRhPct) OR (ABS(fRhPct) > DL_CFW_INF)
   OR (fCoilSurfTempC <> fCoilSurfTempC) OR (ABS(fCoilSurfTempC) > DL_CFW_INF)
   OR (fFrostThreshC <> fFrostThreshC) OR (ABS(fFrostThreshC) > DL_CFW_INF)
   OR (fDpMarginK <> fDpMarginK) OR (ABS(fDpMarginK) > DL_CFW_INF)
   OR (fThawHystK <> fThawHystK) OR (ABS(fThawHystK) > DL_CFW_INF) THEN
    _bCfgBad := TRUE;                    // 非有限归组态非法锁存 / Non-finite folded into the config latch
END_IF
IF (NOT _bCfgBad) AND ((fThawHystK <= DL_CFW_EPS) OR (tFrostDwell <= T#0MS)
   OR (fDpMarginK < DL_CFW_ZERO)) THEN
    _bCfgBad := TRUE;                    // 回差/时间窗/裕度域非法锁存 / Hysteresis, window and margin domains latched
END_IF
IF bReset THEN
    _bCfgBad   := FALSE;                 // 复位清组态锁存 / Reset clears the config latch
    _bCrossBad := FALSE;                 // 复位清交叉锁存 / Reset clears the cross latch
    _bDefrostL := FALSE;                 // 复位清请求锁存 / Reset clears the request latch
END_IF

(*------------------------------------------------------------------------------
 * 段 4｜湿度钳位与露点内联解算（Device 泳道零外部依赖）
 *      Humidity clamp and the inline dew-point solve
 *-----------------------------------------------------------------------------*)
_fRhUse := MIN(MAX(fRhPct, DL_CFW_RH_MIN), DL_CFW_RH_MAX); // 湿度双侧钳位（对数域下限保证） / Two-sided humidity clamp
_fGamma := LN(_fRhUse / 100.0);          // 中间量 ln(RH/100) [无量纲]，恒 <= 0 / Intermediate, always <= 0
_fDpCalc := DL_CFW_MAGNUS_B * _fGamma / (DL_CFW_MAGNUS_A - _fGamma); // Magnus 露点反解 [摄氏度]，分母恒 > 17 / Magnus dew-point solve, denominator always > 17
fDewPointC := _fDpCalc;                  // 露点诊断出口 / Dew-point diagnostics outlet

(*------------------------------------------------------------------------------
 * 段 5｜传感器交叉校验：露点 > 干球 + 容差 → 物理不可能，判通道异常
 *      Sensor cross-check: dew point above the dry bulb is impossible
 *-----------------------------------------------------------------------------*)
IF (NOT _bCfgBad) AND (_fDpCalc > (fAirTempC + DL_CFW_CROSS_K)) THEN
    _bCrossBad := TRUE;                  // 交叉校验失败锁存（安全侧锁存请求） / Cross-check failure latched, request latched on the safe side
    _bDefrostL := TRUE;                  // 安全侧：宁多除一次，不漏霜 / Safe side: defrost rather than miss frost
END_IF

(*------------------------------------------------------------------------------
 * 段 6｜驻留计时无条件刷新（R40：CASE 之外每拍必调）
 *      Dwell timer refreshed unconditionally per R40
 *-----------------------------------------------------------------------------*)
fbDwell(IN := (_eState = E_DL_CoilFrostState.eMonitor)
             AND (fCoilSurfTempC <= fFrostThreshC)
             AND (fCoilSurfTempC <= (_fDpCalc - fDpMarginK)),
        PT := tFrostDwell);              // 双判据驻留窗 / Dual-criteria dwell window

(*------------------------------------------------------------------------------
 * 段 7｜相位机（CASE 含 ELSE 兜底；未使能/异常落故障态）
 *      Phase machine with ELSE fallback
 *-----------------------------------------------------------------------------*)
IF (NOT bEnable) OR _bCfgBad OR _bCrossBad THEN
    _eState := E_DL_CoilFrostState.eFault; // 未使能或异常转故障态 / Not enabled or anomaly, fault
ELSE
CASE _eState OF

    E_DL_CoilFrostState.eIdle:             // 空闲：使能进监视
        IF bEnable THEN
            _eState := E_DL_CoilFrostState.eMonitor; // 进监视 / To monitor
        END_IF

    E_DL_CoilFrostState.eMonitor:          // 监视：双判据驻留满进霜窗
        IF NOT bEnable THEN
            _eState := E_DL_CoilFrostState.eFault; // 使能撤销转故障 / Enable dropped, fault
        ELSIF fbDwell.Q THEN
            _bInfoFrost := TRUE;           // 霜窗确认（信息级，拍 N 进入） / Frost window confirmed, info
            _bDefrostL := TRUE;            // 除霜请求锁存建立 / Defrost request latched
            _eState := E_DL_CoilFrostState.eDefrost; // 进除霜态 / To defrost
        END_IF

    E_DL_CoilFrostState.eFrost:            // 霜窗：请求已锁存，转除霜态保持
        _bDefrostL := TRUE;                // 请求保持 / Request held
        _eState := E_DL_CoilFrostState.eDefrost; // 进除霜态 / To defrost

    E_DL_CoilFrostState.eDefrost:          // 除霜：回差退出或复位解除
        IF (NOT bEnable) OR _bCfgBad THEN
            _eState := E_DL_CoilFrostState.eFault; // 异常转故障 / Anomaly, fault
        ELSIF fCoilSurfTempC > (fFrostThreshC + fThawHystK) THEN
            _bInfoDone := TRUE;            // 除霜完成回差退出（信息级） / Thaw hysteresis exit, info
            _bDefrostL := FALSE;           // 请求解除 / Request released
            _eState := E_DL_CoilFrostState.eMonitor; // 回监视 / Back to monitor
        END_IF

    E_DL_CoilFrostState.eFault:            // 故障：复位沿且原因消失回空闲
        IF bReset AND (NOT _bCfgBad) AND (NOT _bCrossBad) THEN
            _eState := E_DL_CoilFrostState.eIdle; // 回空闲 / Back to idle
        END_IF

    ELSE                                   // 非法状态兜底（R21：CASE 必带 ELSE）
        _bIllegal := TRUE;                 // 标记非法状态 / Flag the illegal state
        _eState   := E_DL_CoilFrostState.eFault; // 回故障态 / Back to fault
END_CASE
END_IF

(*------------------------------------------------------------------------------
 * 段 8｜码位出口与放行（故障级码 3 行内置 bError，R45/R101 配对）
 *      Code outlet and release, fault codes paired with bError
 *-----------------------------------------------------------------------------*)
IF _bIllegal THEN
    eErr   := 16#0003_0362;                // 故障级：状态机兜底 / Fault: state machine fallback
    bError := TRUE;                        // 置故障标志 / Raise the fault flag
ELSIF _bCrossBad THEN
    eErr   := 16#0003_0361;                // 故障级：传感器交叉校验失败 / Fault: sensor cross-check failed
    bError := TRUE;                        // 置故障标志 / Raise the fault flag
ELSIF _bCfgBad THEN
    eErr   := 16#0003_0360;                // 故障级：组态非法 / Fault: illegal configuration
    bError := TRUE;                        // 置故障标志 / Raise the fault flag
ELSIF _bInfoDone THEN
    eErr := 16#0003_018B;                  // 信息级：除霜完成回差退出 / Info: thaw hysteresis exit
ELSIF _bInfoFrost THEN
    eErr := 16#0003_018A;                  // 信息级：结霜窗确认 / Info: frost window confirmed
END_IF

bFrostWindow := (_eState = E_DL_CoilFrostState.eDefrost); // 霜窗电平 = 除霜态（锁存期） / Frost level equals the defrost phase
bDefrostReq  := _bDefrostL;              // 除霜请求出口 = 锁存量（R99） / Defrost request outlet equals the latch
bValid := (NOT bError) AND bEnable AND (_eState <> E_DL_CoilFrostState.eIdle); // 空闲/故障/未使能输出不可用 / Outputs unusable in idle, fault or disabled
eState := _eState;                       // 相位出口 / Phase outlet
END_FUNCTION_BLOCK

(* ---- FB_DL_ColorChangeSeq.st ---- *)
(*
  Name: FB_DL_ColorChangeSeq
  Category: DL_Device
  Version: 1.0.0
  Round: R89 / 2026-11-25
  开源溯源：clean-room 自研（族 涂装喷涂线，ST 开源生态实测 0 命中，无外部代码引入）
  功能：换色清洗顺序：吹扫→溶剂冲洗→再吹干→试喷确认，三段时间与试喷确认窗口各自独立 TON。
  边界条件：① 三段时长必须 > 0，否则组态非法直接锁故障（本件无码出口，成因由相位 + xFault 表达）；
            ② 吹扫/冲洗/吹干各用独立 TON，PT 分别取 tBlowS / tFlushS / tDryS，禁跨相共用（R100）；
            ③ 试喷确认窗为固定时窗 DL_CCS_PILOT（10 s，无外部引脚），超窗未确认即锁故障；
            ④ 完成脉冲两段式：相内只置 _bDone，出口统一映射单拍，避免同拍抹除（R187）；
            ⑤ 故障解除唯一路径：故障相内 xStart 释放（R152），清锁存回 eIdle。
  状态机：eIdle / eBlow / eFlush / eDry / ePilot / eDone / eFault（CASE 含 ELSE 兜底）。
*)
TYPE E_DL_Ccs2Phase :
(
    eIdle  := 0,        (* 待机：等启动沿 / Idle, waiting for start edge *)
    eBlow  := 10,       (* 吹扫相：压缩空气吹除残漆 / Blow phase, purge residual paint *)
    eFlush := 20,       (* 冲洗相：溶剂冲洗管路 / Flush phase, solvent *)
    eDry    := 30,      (* 吹干相：吹干溶剂残留 / Dry phase, air dry *)
    ePilot := 40,       (* 试喷相：等试喷确认 / Pilot spray, waiting confirmation *)
    eDone  := 50,       (* 完成相：保持至启动释放 / Done, holds until start released *)
    eFault := 90        (* 故障相：锁存待释放 / Fault latched, awaiting release *)
);
END_TYPE

FUNCTION_BLOCK FB_DL_ColorChangeSeq
VAR_INPUT
    xStart : BOOL;          (* 启动命令（上升沿起序） [-] Start command, rising edge *)
    tBlowS : TIME;          (* 吹扫时长 [ms] Blow duration [ms] *)
    tFlushS : TIME;         (* 溶剂冲洗时长 [ms] Flush duration [ms] *)
    tDryS : TIME;           (* 吹干时长 [ms] Dry duration [ms] *)
    xPilotOk : BOOL;        (* 试喷确认（膜厚/色差合格） [-] Pilot spray confirmed *)
END_VAR
VAR_OUTPUT
    eState : E_DL_Ccs2Phase;    (* 当前相 [-] Present phase *)
    xValveSolvent : BOOL;       (* 溶剂阀指令（仅冲洗相） [-] Solvent valve command *)
    xValveAir : BOOL;           (* 空气阀指令（吹扫/吹干相） [-] Air valve command *)
    xDone : BOOL;               (* 换色完成单拍脉冲 [-] One-scan done pulse *)
    xFault : BOOL;              (* 故障锁存标志 [-] Fault latched *)
END_VAR
VAR
    _ePhase : E_DL_Ccs2Phase := E_DL_Ccs2Phase.eIdle;  (* 内部相（CASE 唯一写入目标） [-] Internal phase *)
    _bDone : BOOL := FALSE;         (* 单拍完成标志（段 1 预清） [-] One-scan done flag *)
    _bFaultLatch : BOOL := FALSE;   (* 故障锁存位 [-] Fault latch *)
    _bReqFault : BOOL := FALSE;     (* 单拍故障请求（段 1 预清） [-] Fault request *)
    tonBlow : TON;                  (* 吹扫计时（段 0 无条件调用） / Blow timer *)
    tonFlush : TON;                 (* 冲洗计时（段 0 无条件调用） / Flush timer *)
    tonDry : TON;                   (* 吹干计时（段 0 无条件调用） / Dry timer *)
    tonPilot : TON;                 (* 试喷确认窗（段 0 无条件调用） / Pilot confirm window *)
    rtStart : R_TRIG;               (* 启动沿（段 0 无条件调用） / Start edge *)
END_VAR
VAR CONSTANT
    DL_CCS2_PILOT : TIME := T#10S;  (* 试喷确认窗（固定时窗） [ms] Pilot confirmation window [ms] *)
END_VAR
(* —— 段 0：沿与四 TON 无条件周期刷新（R7），IN 仅由相位派生 —— *)
rtStart(CLK := xStart);                                                 (* 启动沿 / Start edge *)
tonBlow(IN := (_ePhase = E_DL_Ccs2Phase.eBlow), PT := tBlowS);          (* 吹扫计时 / Blow timer *)
tonFlush(IN := (_ePhase = E_DL_Ccs2Phase.eFlush), PT := tFlushS);       (* 冲洗计时 / Flush timer *)
tonDry(IN := (_ePhase = E_DL_Ccs2Phase.eDry), PT := tDryS);             (* 吹干计时 / Dry timer *)
tonPilot(IN := (_ePhase = E_DL_Ccs2Phase.ePilot), PT := DL_CCS2_PILOT); (* 试喷窗 / Pilot window *)
(* —— 段 1：单拍量预清 + 组态故障请求 —— *)
_bDone := FALSE;
_bReqFault := FALSE;
IF (tBlowS <= T#0S) OR (tFlushS <= T#0S) OR (tDryS <= T#0S) THEN
    _bReqFault := TRUE;                         (* 组态非法：时长为零 / Configuration bad, zero duration *)
END_IF
(* —— 段 2：故障锁存解除（唯一路径 = 故障相内 xStart 释放，R152） —— *)
IF _bFaultLatch AND (NOT xStart) THEN
    _bFaultLatch := FALSE;                      (* 清锁存 / Clear latch *)
    _ePhase := E_DL_Ccs2Phase.eIdle;            (* 迁回待机 / Back to idle *)
END_IF
(* —— 段 3：主状态机（ENUM + CASE，ELSE 兜底） —— *)
CASE _ePhase OF
E_DL_Ccs2Phase.eIdle:
    IF rtStart.Q AND (NOT _bFaultLatch) THEN
        _ePhase := E_DL_Ccs2Phase.eBlow;        (* 起序 → 吹扫 / Start, blow *)
    END_IF
E_DL_Ccs2Phase.eBlow:
    IF tonBlow.Q THEN
        _ePhase := E_DL_Ccs2Phase.eFlush;       (* 吹扫到时 → 冲洗 / Blow done, flush *)
    END_IF
E_DL_Ccs2Phase.eFlush:
    IF tonFlush.Q THEN
        _ePhase := E_DL_Ccs2Phase.eDry;         (* 冲洗到时 → 吹干 / Flush done, dry *)
    END_IF
E_DL_Ccs2Phase.eDry:
    IF tonDry.Q THEN
        _ePhase := E_DL_Ccs2Phase.ePilot;       (* 吹干到时 → 试喷 / Dry done, pilot *)
    END_IF
E_DL_Ccs2Phase.ePilot:
    IF xPilotOk THEN
        _bDone := TRUE;                         (* 单拍完成（段 1 预清） / One-scan done *)
        _ePhase := E_DL_Ccs2Phase.eDone;        (* → 完成相 / To done *)
    ELSIF tonPilot.Q THEN
        _bReqFault := TRUE;                     (* 试喷窗超时未确认 / Pilot window expired *)
    END_IF
E_DL_Ccs2Phase.eDone:
    IF NOT xStart THEN
        _ePhase := E_DL_Ccs2Phase.eIdle;        (* 启动释放 → 待机 / Start released, idle *)
    END_IF
E_DL_Ccs2Phase.eFault:
    _bReqFault := FALSE;                        (* 故障相驻留：锁存已置，不再新发请求 *)
ELSE
    _bReqFault := TRUE;                         (* 非法相兜底 / Illegal phase fallback *)
END_CASE
(* —— 段 4：故障请求统一落地（唯一锁存点 + 同步迁相，R187/R252） —— *)
IF _bReqFault AND (NOT _bFaultLatch) THEN
    _bFaultLatch := TRUE;                       (* 锁存 / Latch *)
    _ePhase := E_DL_Ccs2Phase.eFault;           (* 同步迁相 / Migrate to fault *)
END_IF
(* —— 段 5：统一出口（各出口单点赋值） —— *)
eState := _ePhase;
xValveSolvent := (_ePhase = E_DL_Ccs2Phase.eFlush) AND (NOT _bFaultLatch);
xValveAir := ((_ePhase = E_DL_Ccs2Phase.eBlow) OR (_ePhase = E_DL_Ccs2Phase.eDry)) AND (NOT _bFaultLatch);
xDone := _bDone;
xFault := _bFaultLatch;
END_FUNCTION_BLOCK
